(* IEC 61131-3 sources: IRIS-Project/LASAL CONTROL SOFTWARE/LasalProject_2025_09_12/Runtime/%LASALAPPDATA%/Runtime/Library/Loader/Source/code (part 9) *)

END_FUNCTION

//------------------------------------------------------------------------------
// RecvBuf
//
//  This function reads data from a connection. The data is buffered. A tcp-recv
//  operation receives as much data as possible into the internal rx buffer.
//  Data that is not needed by the caller remains in the internal rx buffer.
//  This techniqe is used to avoid multiple small reads from the tcp/ip
//  connection.
//
// Return value
//  If the function succeeds, the return value is the number of bytes read,
//  otherwise a tcp-user error code is returned.
//------------------------------------------------------------------------------
FUNCTION RecvBuf
VAR_INPUT
    bsock         : ^bufferedSocket;
    buf           : ^CHAR;
    len           : UDINT;
    timeout_ms    : UDINT;      // timeout, in milliseconds
END_VAR
VAR_OUTPUT
    retval        : DINT;
END_VAR
VAR
    reqMsg        : msgNopReq;
END_VAR

  #ifdef DEBUG
  ChkBuffer(bsock);
  #endif

  IF bsock^.bytesInRxBuf = 0 THEN
    // The receive buffer is empty

    // Receive as much as possible into the rx buffer
    retval := OS_TCP_USER_RECV(bsock^.sock,
                               #bsock^.rxBuf[0],
                               bsock^.sizeOfRxBuf,
                               0,
                               timeout_ms
                               );
    IF retval <= 0 THEN
#ifdef DEBUG
      IF (retval <> TCP_NOT_READY) | (timeout_ms > 0) THEN
        DEBUGLOG2("%010d-OS_TCP_USER_RECV(sock %d) failed, rc=%d", TO_UDINT(bsock^.sock), TO_UDINT(retval));
      END_IF;
#endif
      IF retval <> TCP_NOT_READY THEN
        CloseBufferedSock(bsock);
      END_IF;
      RETURN;
    END_IF;
    bsock^.bytesInRxBuf += TO_UDINT(retval);
    DEBUG_VERBOSE3("%010d-OS_TCP_USER_RECV(sock %d): %d bytes received, new bytesInRxBuf=%d", TO_UDINT(bsock^.sock), TO_UDINT(retval), TO_UDINT(bsock^.bytesInRxBuf));

    IF bsock^.fAckRcvdData THEN
      // send something after data received to avoid delayed ack
      IF bsock^.bytesInTxBuf > 0 THEN
        FLUSH_TXBUF(bsock);
      ELSE
        SendCmdMsg(bsock,
                   CMD_NOP,
                   0,                 // Type and Ack field of command (type: request, ack: no response is required)
                   #reqMsg$cMessage,
                   SIZEOF(reqMsg),
                   0,                 // timeout: 5 sec.
                   1,                 // use buffered sends
                   1                  // fFlush
                  );
      END_IF;
    END_IF;

  END_IF; // empty rx buffer

  // copy data from the buffer to the caller
  IF len < bsock^.bytesInRxBuf THEN
    retval := len$DINT;
  ELSE
    retval := bsock^.bytesInRxBuf$DINT;
  END_IF;
  IF buf <> NIL THEN
    _memcpy(buf, #bsock^.rxBuf[bsock^.rxBufStrtInd], TO_UDINT(retval));
  END_IF;

  // adjust buffer variables
  bsock^.bytesInRxBuf -= TO_UDINT(retval);
  bsock^.rxBufStrtInd += TO_UDINT(retval);
  IF bsock^.bytesInRxBuf = 0 THEN
    bsock^.rxBufStrtInd := 0;
  END_IF;

  #ifdef DEBUG
  ChkBuffer(bsock);
  #endif

END_FUNCTION

//------------------------------------------------------------------------------
// UnRecvBuf
//
//  This function places len bytes back into the internal rx buffer.
//
// Return value
//  The number of bytes placed into the buffer.
//------------------------------------------------------------------------------
FUNCTION UnRecvBuf
VAR_INPUT
    bsock          : ^bufferedSocket;
    buf            : ^CHAR;
    len            : UDINT;
END_VAR
VAR_OUTPUT
    retval         : UDINT;
END_VAR
VAR
    bytesFree      : UDINT;    // total number of free bytes in the rx buffer
END_VAR

  #ifdef DEBUG
  ChkBuffer(bsock);
  #endif

  bytesFree      := bsock^.sizeOfRxBuf - bsock^.bytesInRxBuf;

  IF len < bytesFree THEN
    retval := len;
  ELSE
    retval := bytesFree;
  END_IF;

  IF retval > bsock^.rxBufStrtInd THEN
    // move the data in rxBuf to the end of the buffer
    _memmove(#bsock^.rxBuf[retval], #bsock^.rxBuf[bsock^.rxBufStrtInd], bsock^.bytesInRxBuf);
    bsock^.rxBufStrtInd := retval;
  END_IF;

  bsock^.rxBufStrtInd -= retval;
  bsock^.bytesInRxBuf += retval;
  _memcpy(#bsock^.rxBuf[bsock^.rxBufStrtInd], buf, retval);

  #ifdef DEBUG
  ChkBuffer(bsock);
  #endif

END_FUNCTION

//------------------------------------------------------------------------------
// ReadN
//
//  This function reads n bytes from a connection.
//
// Return value
//  If the function succeeds, the return value is the number of bytes requested,
//  otherwise a tcp-user error code is returned.
//------------------------------------------------------------------------------
FUNCTION ReadN
VAR_INPUT
    bsock         : ^bufferedSocket;
    buf           : ^CHAR;
    len           : UDINT;
    timeout_ms    : UDINT;      // timeout, in milliseconds
END_VAR
VAR_OUTPUT
    retval        : DINT;
END_VAR
VAR
    ptr           : ^CHAR;
    bytesToRead   : UDINT;      // number of bytes to read
    bytesRead     : UDINT;      // number of bytes already read
END_VAR

    bytesToRead := len;
    bytesRead   := 0;
    ptr         := buf;
    WHILE bytesToRead > 0 DO
      retval := RecvBuf(bsock, ptr, bytesToRead, timeout_ms);
      IF retval <= 0 THEN
        // In the case of an error place already read data back to the buffer
        IF UnRecvBuf(bsock, buf, bytesRead) <> bytesRead THEN
          // This code should never be reached !
          DEBUGLOG1("%010d-ReadN(sock %d): UnRecvBuf failed", TO_UDINT(bsock^.sock));
          CloseBufferedSock(bsock);
          retval := ERR_CONN_BROKEN;
        END_IF;
        RETURN;
      END_IF;
      bytesToRead -= retval$UDINT;
      bytesRead   += retval$UDINT;
      ptr         += retval;
    END_WHILE;

    retval := bytesRead$DINT;

END_FUNCTION

//------------------------------------------------------------------------------
// ReadVRec
//
//  This function reads a record with a variable length.
//
// Return value
//  If the function succeeds, the return value is the number of bytes received
//  in the data field (without vrec-header).
//
// Remarks
//  When the size of the buffer is too small for the message, the connection is
//  closed.
//------------------------------------------------------------------------------
FUNCTION ReadVRec
VAR_INPUT
    bsock         : ^bufferedSocket;
    vrec          : ^vRecord;    // the variable record buffer
    len           : UDINT;      // length of the buffer incl. header
    timeout_ms    : UDINT;      // timeout, in milliseconds
END_VAR
VAR_OUTPUT
    retval        : DINT;
END_VAR

  // first read the vrec-header
  retval := ReadN(bsock, (#vrec^.vHdr)$^CHAR, SIZEOF(vrec^.vHdr), timeout_ms);
  IF retval <= 0 THEN
    RETURN;
  END_IF;

  // check if the header is valid
  IF vrec^.vHdr.id <> 0xFACE THEN
    DEBUGLOG1("%010d-ReadVRec(sock %d): invalid vrec-hdr received", TO_UDINT(bsock^.sock));
    CloseBufferedSock(bsock);
    retval := ERR_INVALID_VRECHDR;
    RETURN;
  END_IF;

  // check how many data fits into the buffer
  IF (vrec^.vHdr.dataLen + SIZEOF(vrec^.vHdr)) > len THEN
    DEBUGLOG1("%010d-ReadVRec(sock %d): buffer too small", TO_UDINT(bsock^.sock));
    CloseBufferedSock(bsock);
    retval := ERR_BUF_TOO_SMALL;
    RETURN;
  END_IF;

  // read the data of the variale record
  retval := ReadN(bsock, (#vrec^.data)$^CHAR, vrec^.vHdr.dataLen, timeout_ms);
  IF retval <= 0 THEN
    // error: write the vrec-header back to the buffer
    IF UnRecvBuf(bsock, (#vrec^.vHdr)$^CHAR, SIZEOF(vrec^.vHdr)) <> SIZEOF(vrec^.vHdr) THEN
      // This code should never be reached !
      DEBUGLOG1("%010d-ReadVRec(sock %d): UnRecvBuf failed", TO_UDINT(bsock^.sock));
      CloseBufferedSock(bsock);
      retval := ERR_CONN_BROKEN;
    END_IF;
    RETURN;
  END_IF;

END_FUNCTION

//------------------------------------------------------------------------------
// ReadCmdMsg
//
//  This function reads a command message.
//
// Return value
//  If the function succeeds, the return value is the number of bytes received
//  in the data field (without vrec-header).
//
// Remarks
//  When the size of the buffer is too small for the message, the rest of the
//  message received and discarded.
//------------------------------------------------------------------------------
FUNCTION ReadCmdMsg
VAR_INPUT
    bsock         : ^bufferedSocket;
    msg           :^cMessage;   // the message
    len           : UDINT;      // length of the message incl. header
    timeout_ms    : UDINT;      // timeout, in milliseconds
    ack           :^UDINT;      // acknowledge field received (optional)
    cmd           : UDINT;      // matching command of the message (n/a for requests)
    typeMask      : UDINT;      // specifies which type (req.,resp.or both) is expected
END_VAR
VAR_OUTPUT
    retval        : DINT;
END_VAR

  retval := ReadVRec(bsock, msg$^vRecord, len, timeout_ms);
  IF retval <= 0 THEN
    RETURN;
  END_IF;

  IF retval < SIZEOF(msg^.cHdr.cmd) THEN
    // at least the header must be available
    DEBUGLOG1("%010d-ReadCmdMsg(sock %d): missing cmd-hdr", TO_UDINT(bsock^.sock));
    CloseBufferedSock(bsock);
    retval := ERR_INVALID_CMSGHDR;
    RETURN;
  END_IF;

  // check if the type of message is expected by the caller
  IF msg^.cHdr.cmd AND MASK_CMD_ISRESP THEN
     // a response is received

    IF (typeMask AND CMD_TYPE_RESP) = 0 THEN
      DEBUGLOG1("%010d-ReadCmdMsg(sock %d): unexpected resonse received", TO_UDINT(bsock^.sock));
      CloseBufferedSock(bsock);
      retval := ERR_INVALID_CMSGTYPE;
    END_IF;
    IF (msg^.cHdr.cmd AND MASK_CMD_CODE) <> cmd THEN
      DEBUGLOG1("%010d-ReadCmdMsg(sock %d): cmd-code in response does not match", TO_UDINT(bsock^.sock));
      CloseBufferedSock(bsock);
      retval := ERR_INVALID_CMSGCODE;
    END_IF;
    IF (msg^.cHdr.cmd AND MASK_CMD_ACK) = 0 THEN
      DEBUGLOG1("%010d-ReadCmdMsg(sock %d): nack received", TO_UDINT(bsock^.sock));
      CloseBufferedSock(bsock);
      retval := ERR_NACK_RECEIVED;
    END_IF;

  ELSE
    // a request is received

    IF (typeMask AND CMD_TYPE_REQ) = 0 THEN
      DEBUGLOG1("%010d-ReadCmdMsg(sock %d): unexpected request received", TO_UDINT(bsock^.sock));
      CloseBufferedSock(bsock);
      retval := ERR_INVALID_CMSGTYPE;
    END_IF;

  END_IF;

  // extract the ack field
  IF ack <> NIL THEN
    ack^ := msg^.cHdr.cmd AND MASK_CMD_ACK;
  END_IF;

END_FUNCTION

//------------------------------------------------------------------------------
// UpdateCell
//
// Return value:
//  Error                                                     : <=0
//  When udLastUpdate did not expire                          : 1
//  When udLastUpdate expired, but dData did not change       : 2
//  When udLastUpdate expired, and dData changed (transfer)   : 3
//------------------------------------------------------------------------------
#ifdef COMLINK_TCP_SERVER
FUNCTION UpdateCell
VAR_INPUT
    pRefrConn     : ^refrConnBlock;
    pUpdCell      : ^comStCell;  // pointer to cell in updatelist
    iOff          : UINT;
END_VAR
VAR_OUTPUT
    retval        : DINT;
END_VAR
VAR
    reqMsg        : msgUpdCellReq; // request structure for command CMD_UPDCELL
    dData         : DINT;
    rc            : DINT;
END_VAR

  retval := 1;

  if( pUpdCell = NIL )then
    return;
  end_if;

  IF pRefrConn^.bsock.fTxBufferShortage <> 0 THEN
    // in the case of a buffer shortage do not send any updatecells
    RETURN;
  END_IF;

  IF QUERY_FREE_TXBUF(pRefrConn^.bsock) < (2 * SIZEOF(reqMsg)) THEN
    // when there is no more space for 2 messages, then enter buffer shortage
    DEBUGLOG0("%010d-UpdateCell: entering tx buffer shortage");
    pRefrConn^.bsock.fTxBufferShortage := 1;
    // try to send all unsent data
    FLUSH_TXBUF(#pRefrConn^.bsock);
  END_IF;

  IF (ops.tAbsolute - pUpdCell^.udLastUpdate) < (pUpdCell^.udUpdateRate AND 16#FFFF) THEN
    // udLastUpdate did not expire
    RETURN;
  END_IF;

  IF pUpdCell^.pCh = NIL THEN
    RETURN;
  END_IF;

  retval := 2;

  IF (pUpdCell^.udUpdateRate and UPDRATE_FLAG_IS_VBI) THEN
    dData := (pUpdCell^.pCh$^virtualBaseInit^.getCrc())$DINT;
  ELSIF (pUpdCell^.udUpdateRate AND UPDRATE_FLAG_IS_MERKEREX) THEN
     dData := (pUpdCell^.pCh$^merkerex^.getcrc())$DINT;
  ELSIF (pUpdCell^.udUpdateRate AND UPDRATE_FLAG_IS_GLOBALVAR) THEN
//    dData := (pUpdCell^.pCh$^DINT)^;
    dData := UpDateGlobalVar(pUpdCell^.pCh, pUpdCell^.udUpdateRate);
  ELSE
    dData := rd(pUpdCell^.pCh);
  END_IF;

  IF dData = pUpdCell^.dData & (pUpdCell^.udUpdateRate and UPDRATE_FLAG_FORCE_CHANGE) = 0 THEN
    // dData did not change
    pUpdCell^.udLastUpdate := ops.tAbsolute;
    RETURN;
  END_IF;
  pUpdCell^.udUpdateRate := pUpdCell^.udUpdateRate AND NOT UPDRATE_FLAG_FORCE_CHANGE;

  retval := 3;

  // prepare the request message structure
  reqMsg.iOff  := iOff;
  reqMsg.pCh   := pUpdCell^.pCh;
  reqMsg.dData := dData;

  // Send the request
  rc := SendCmdMsg(#pRefrConn^.bsock,
                   CMD_UPDCELL,
                   0,                // Type and Ack field of command (type: request, ack: no response required)
                   #reqMsg$cMessage,
                   SIZEOF(reqMsg),
                   0,                // timeout: non-blocking
                   1,                // use buffered sends
                   pRefrConn^.bsock.fTxBufferShortage // fFlush
                  );
  IF rc <= 0 THEN
    DEBUGLOG2("%010d-*** UpdateCell(VarPos %d): SendCmdMsg failed, rc=%d", TO_UDINT(iOff), TO_UDINT(rc));
    retval := rc;
  ELSE
    //DEBUGLOG3("%010d-UpdateCell: UPDCELL request sent, conn=0x%08X, VarPos=%d, dData=0x%08X", pRefrConn$UDINT, TO_UDINT(iOff), TO_UDINT(dData));
    pUpdCell^.dData := dData;
    pUpdCell^.udLastUpdate := ops.tAbsolute;
  END_IF;

END_FUNCTION
#endif

//------------------------------------------------------------------------------
// UpdateListProcessor
//------------------------------------------------------------------------------
#ifdef COMLINK_TCP_SERVER
FUNCTION UpdateListProcessor
VAR_INPUT
    pRefrConn     : ^refrConnBlock;
END_VAR
VAR
    list          : ^updateList;
    pUpdCell      : ^comStCell;  // pointer to cell in updatelist
    pStrtCell     : ^comStCell;
END_VAR

  if( pRefrConn = NIL )then
    return;
  end_if;
  if( pRefrConn^.ptr = NIL )then
    return;
  end_if;
  list := #pRefrConn^.ptr^.statList;
  if( list = NIL )then
    return;
  end_if;

  IF list^.nbrRefrCells > 0 THEN
    pStrtCell := list^.pActCell;
    WHILE 1 DO
      pUpdCell := list^.pActCell;

      UpdateCell(pRefrConn, pUpdCell, list^.actInd$UINT);
      IF pRefrConn^.bsock.sock < 0 THEN
        RETURN;
      END_IF;

      IF (list^.actInd + 1) >= list^.nbrRefrCells THEN
        list^.actInd   := 0;
        list^.pActCell := list^.pFirstCell;
      ELSE
        list^.actInd   += 1;
        list^.pActCell += SIZEOF(list^.pActCell^);
      END_IF;

      IF pStrtCell = list^.pActCell THEN
        EXIT;
      END_IF;
    END_WHILE;
  END_IF;

  list := #pRefrConn^.ptr^.dynList;
  if( list = NIL )then
    return;
  end_if;
  IF list^.nbrRefrCells > 0 THEN
    pStrtCell := list^.pActCell;
    WHILE 1 DO
      pUpdCell := list^.pActCell;

      if( pUpdCell = NIL )then
        return;
      end_if;
      UpdateCell(pRefrConn, pUpdCell, (list^.actInd + 1000)$UINT);
      IF pRefrConn^.bsock.sock < 0 THEN
        RETURN;
      END_IF;

      IF (list^.actInd + 1) >= list^.nbrRefrCells THEN
        list^.actInd   := 0;
        list^.pActCell := list^.pFirstCell;
      ELSE
        list^.actInd   += 1;
        list^.pActCell += SIZEOF(list^.pActCell^);
      END_IF;

      IF pStrtCell = list^.pActCell THEN
        EXIT;
      END_IF;
    END_WHILE;
  END_IF;

END_FUNCTION
#endif

//------------------------------------------------------------------------------
// SendAliveMessage_TCP
//------------------------------------------------------------------------------
#ifdef COMLINK_TCP_SERVER
FUNCTION SendAliveMessage_TCP
VAR_INPUT
    pRefrConn     : ^refrConnBlock;
END_VAR
VAR_OUTPUT
    retval        : DINT;
END_VAR
VAR
    reqMsg        : msgIamAliveReq; // request structure for command CMD_UPDCELL
    rc            : DINT;
END_VAR

  retval := 1;

  IF pRefrConn^.bsock.fTxBufferShortage <> 0 THEN
    // in the case of a buffer shortage do not send any requests
    RETURN;
  END_IF;

  IF QUERY_FREE_TXBUF(pRefrConn^.bsock) < (2 * SIZEOF(reqMsg)) THEN
    // when there is no more space for 2 messages, then enter buffer shortage
    DEBUGLOG0("%010d-SendAliveMessage_TCP: entering tx buffer shortage");
    pRefrConn^.bsock.fTxBufferShortage := 1;
    // try to send all unsent data
    FLUSH_TXBUF(#pRefrConn^.bsock);
  END_IF;

  // Send the request
  rc := SendCmdMsg(#pRefrConn^.bsock,
                   CMD_IAMALIVE,
                   0,                // Type and Ack field of command (type: request, ack: no response required)
                   #reqMsg$cMessage,
                   SIZEOF(reqMsg),
                   0,                // timeout: non-blocking
                   1,                // use buffered sends
                   1                 // fFlush
                  );
  IF rc <= 0 THEN
    DEBUGLOG1("%010d-*** SendAliveMessage_TCP: SendCmdMsg failed, rc=%d", TO_UDINT(rc));
    retval := rc;
  ELSE
    DEBUG_VERBOSE1("%010d-SendAliveMessage_TCP: IAMALIVEL request sent, conn=0x%08X", pRefrConn$UDINT);
  END_IF;
END_FUNCTION
#endif

//------------------------------------------------------------------------------
// SyncRefListsTcp  - siehe Beschreibung von SyncRefLists
//------------------------------------------------------------------------------
#ifdef COMLINK_TCP_SERVER
FUNCTION SyncRefListsTcp
VAR_INPUT
    pCmdConn    : ^cmdConnBlock;
END_VAR
VAR
    obj         : pVoid;
    pHead       : ^IprHead;
    instr       : ^instruct;
    pRefrConn   : ^refrConnBlock;
END_VAR

    pRefrConn := pRefrConnRoot;
    WHILE pRefrConn <> NIL DO
        IF pRefrConn^.ipAddrPeer = pCmdConn^.ipAddrPeer THEN

#ifndef DUMMY_LOADER
            pHead := pCmdConn^.ptr^.com.GetHead();
#endif
            instr := pHead^.pCode;

            IF instr^.opCode = I_WRITE THEN

                obj := instr^.aPara[0]$^pVoid;

                // statische Refresh-Liste durchsuchen
                InvalidateRefListEntry(pRefrConn^.ptr^.statList.pFirstCell, pRefrConn^.ptr^.statList.nbrRefrCells$UINT, obj);

                // dynamische Refresh-Liste durchsuchen
                InvalidateRefListEntry(pRefrConn^.ptr^.dynList.pFirstCell, pRefrConn^.ptr^.dynList.nbrRefrCells$UINT, obj);

            END_IF;

        END_IF;
        pRefrConn := pRefrConn^.next;
    END_WHILE;

END_FUNCTION

FUNCTION GLOBAL SyncRefListsTcpAll
  VAR_INPUT
    lasalid : udint;
  END_VAR
  var
    pRefrConn   : ^refrConnBlock;
  end_var

  pRefrConn := pRefrConnRoot;

  while(pRefrConn <> NIL) do
    // statische Refresh-Liste durchsuchen
    InvalidateRefListEntry(pRefrConn^.ptr^.statList.pFirstCell, pRefrConn^.ptr^.statList.nbrRefrCells$UINT, lasalid$^void);

    // dynamische Refresh-Liste durchsuchen
    InvalidateRefListEntry(pRefrConn^.ptr^.dynList.pFirstCell, pRefrConn^.ptr^.dynList.nbrRefrCells$UINT, lasalid$^void);
    pRefrConn := pRefrConn^.next;
  end_while;

END_FUNCTION
#endif

//------------------------------------------------------------------------------
// Entfernt unbenutzte Verbindungen.
// Es werden alle Verbindungen mit einer bestimmten Remote-IP-Adresse untersucht.
// Wenn die Inst-ID nicht mit der angegebenen übereinstimmt, dann kann es sich
// nur um einen Neustart der Station mit dieser IP-Adresse handeln, da die
// Inst-ID beim Comlink-Init immer neu vergeben wird.
//
// Verbindungen, bei denen die Inst-ID für eine längere Zeit 0 ist, werden
// ebenfalls beendet. Hier handelt es sich um Verbindungen, bei denen abgesteckt
// wurde, bevor CMD_SESSINFO empfangen worden ist.
//
// ApplicationID:
// Wird nur von Comlink Verbindungen von PC-Anwendungen verwendet.
// Wenn auf einem PC mehrere Anwendungen eine Comlink Verbindung verwenden,
// dann kann jede Anwendung eine eigene ApplicationID mitschicken. Damit wird
// verhindert, dass die zweite Anwendung die Verbindung der ersten löscht.
//------------------------------------------------------------------------------
#ifdef COMLINK_TCP_SERVER
FUNCTION DeleteUnusedConnections
VAR_INPUT
    ipAddrPeer   : UDINT;
    instIdOfPeer : UDINT;
    ApplicationID : UDINT;  // ApplicationID
END_VAR
VAR
    pCmdConn   : ^cmdConnBlock;
    pRefrConn   : ^refrConnBlock;
    pCmdConn_next   : ^cmdConnBlock;
    pRefrConn_next  : ^refrConnBlock;
END_VAR

    pCmdConn := pCmdConnRoot;
    WHILE pCmdConn <> NIL DO
        pCmdConn_next := pCmdConn^.next;
        IF ((pCmdConn^.ipAddrPeer = ipAddrPeer) &
            (pCmdConn^.ptr^.instIdOfPeer <> 0) &
            (pCmdConn^.ptr^.instIdOfPeer <> instIdOfPeer) &
            (pCmdConn^.ApplicationID = ApplicationID))
            |
           ((pCmdConn^.ptr^.instIdOfPeer = 0) &
            ((ops.tAbsolute - pCmdConn^.connectTime) > 5000)) THEN
            DEBUGLOG1("%010d-  =====  unused Cmd conn.data block found (ip 08%X) -> releasing block  =====", ipAddrPeer);
            ReleaseConnBlock(TYPE_CMD_CONN, pCmdConn$^connBlock, 0);
            pCmdConn := NIL;
        END_IF;
        pCmdConn := pCmdConn_next;
    END_WHILE;

    pRefrConn := pRefrConnRoot;
    WHILE pRefrConn <> NIL DO
        pRefrConn_next := pRefrConn^.next;
        IF ((pRefrConn^.ipAddrPeer = ipAddrPeer) &
            (pRefrConn^.ptr^.instIdOfPeer <> 0) &
            (pRefrConn^.ptr^.instIdOfPeer <> instIdOfPeer) &
            (pRefrConn^.ApplicationID = ApplicationID))
            |
           ((pRefrConn^.ptr^.instIdOfPeer = 0) &
            ((ops.tAbsolute - pRefrConn^.connectTime) > 5000)) THEN
            DEBUGLOG1("%010d-  =====  unused Refr conn.data block found (ip 08%X) -> releasing block  =====", ipAddrPeer);
            ReleaseConnBlock(TYPE_REFR_CONN, pRefrConn$^connBlock, 0);
            pRefrConn := NIL;
        END_IF;
        pRefrConn := pRefrConn_next;
    END_WHILE;

END_FUNCTION
#endif

//------------------------------------------------------------------------------
// DeleteUnusedRecycleData
//
//  Es werden unbenutzte refresh-connection-data-block's im recycle pool
//  gesucht und wenn gefunden, dann freigegeben.
//
//  Kriterium, ob ein data-block unbenutzt ist:
//  - IP Adresse muss übereinstimmen
//  - InstanceId muss vorhanden, aber unterschiedlich sein
//  - ApplicationID muss übereinstimmen
//------------------------------------------------------------------------------
#ifdef COMLINK_TCP_SERVER
FUNCTION DeleteUnusedRecycleData
VAR_INPUT
    ipAddrPeer   : UDINT;
    instIdOfPeer : UDINT;
    ApplicationID : UDINT;  // ApplicationID
END_VAR
VAR
    pDataWork : ^refrConnData;
    pDataPrev : ^refrConnData;
END_VAR

  pDataPrev := NIL;
  pDataWork := pRefrConnDataRoot;
  WHILE pDataWork <> NIL DO
    IF ((pDataWork^.ipAddrPeer = ipAddrPeer) &
        (pDataWork^.instIdOfPeer <> 0) &
        (pDataWork^.instIdOfPeer <> instIdOfPeer) &
        (pDataWork^.ApplicationID = ApplicationID)) THEN
      // remove it from the recycle pool
      IF pDataPrev = NIL THEN
        pRefrConnDataRoot  := pDataWork^.next;
      ELSE
        pDataPrev^.next := pDataWork^.next;
      END_IF;
      DEBUGLOG1("%010d-  =====  unused recycle refr conn.data block found (ip 08%X) -> releasing block  =====", ipAddrPeer);
      FreeRefrConnData(pDataWork);
      nbrRecycled -= 1;
      EXIT;
    END_IF;
    pDataPrev := pDataWork;
    if( pDataWork = pDataWork^.next )then
      exit;
    end_if;
    pDataWork := pDataWork^.next;
  END_WHILE;

END_FUNCTION
#endif

//------------------------------------------------------------------------------
// CmdMsgListener
//
//  This function serves incoming requests from the client on the command
//  channel.
//------------------------------------------------------------------------------
#ifdef COMLINK_TCP_SERVER
FUNCTION CmdMsgListener
VAR_INPUT
    pCmdConn         : ^cmdConnBlock;
END_VAR
VAR_OUTPUT
    retval    : DINT;
END_VAR
VAR
    cmsg      : cMessage512;
    ackRcvd   : UDINT;        // received ack-field
    ackSend   : UDINT;        // ack-field to send
    dataLen   : UDINT;
    bNext     : UDINT;
    msgLen    : UDINT;
    pResu     : ^results;
    cmd       : UDINT;
    pCmdConnTemp : ^cmdConnBlock;
    rc : DINT;
    releaseFlag : UDINT;
END_VAR

  retval := 0;
  releaseFlag := 0;

  #ifdef LOADER_TCP_MODERATE
    if (pCmdConn^.bsock.isDataAvailable = false) then
      return;
    end_if;
  #endif

  rc := ReadCmdMsg(#pCmdConn^.bsock,
                       #cmsg$cMessage,
                       sizeof(cmsg),
                       0,                   // timeout: 0 means non blocking
                       #ackRcvd,            // received ack field
                       0,                   // matching cmd-code (n/a for requests)
                       CMD_TYPE_REQ         // accept only request types
                      );
  IF rc <= 0 THEN
#ifdef DEBUG
    IF rc <> TCP_NOT_READY THEN
      DEBUGLOG2("%010d-*** CmdMsgListener(sock %d): ReadCmdMsg failed, rc=%d", TO_UDINT(pCmdConn^.bsock.sock), TO_UDINT(rc));
    END_IF;
#endif
    RETURN;
  END_IF;

  retval := 1;

  dataLen := cmsg.cHdr.vHdr.dataLen - SIZEOF(cmsg.cHdr.cmd);
  ackSend := 0; // unsupported command
  msgLen  := SIZEOF(cmsg.cHdr);

  cmd := cmsg.cHdr.cmd AND MASK_CMD_CODE;
  CASE cmd OF

    CMD_BEFIPR:
      DEBUG_VERBOSE2("%010d-CmdMsgListener: sock %d - BEFIPR received, dataLen=%d", TO_UDINT(pCmdConn^.bsock.sock), dataLen$UDINT);
      // req-data:
      //    workState   : iprStates;
      //    instr       : instruct;
      // resp-data:
      //    workState   : iprStates;
      //    resu        : results;

      IF (dataLen < SIZEOF(iprStates)) | ((dataLen - SIZEOF(iprStates)) > SIZEOF(instruct)) THEN
        cmsg$msgBefiprResp.workstate := ERROR;
      ELSE
        // execute befipr
#ifndef DUMMY_LOADER
#ifdef LOADER_4_LASAL2
        _memcpy(pCmdConn^.ptr^.com._m.head.pCode, #cmsg$msgBefiprReq.instr, dataLen - SIZEOF(iprStates));
        pCmdConn^.ptr^.com._m.head.workstate := cmsg$msgBefiprReq.workstate;
        pCmdConn^.ptr^.com._m.head.funkSt    := READY;
        pCmdConn^.ptr^.Com._m.resu.uilng :=0;
#else
        _memcpy(pCmdConn^.ptr^.com.head.pCode, #cmsg$msgBefiprReq.instr, dataLen - SIZEOF(iprStates));
        pCmdConn^.ptr^.com.head.workstate := cmsg$msgBefiprReq.workstate;
        pCmdConn^.ptr^.com.head.funkSt    := READY;
        pCmdConn^.ptr^.Com.resu.uilng :=0;
#endif
        cmsg$msgBefiprResp.workstate := pCmdConn^.ptr^.com.BEFIPR(#bNext);
#endif
        SyncRefListsTcp(pCmdConn);
      END_IF;

      // prepare the response
      ackSend := MASK_CMD_ACK;  // command processed
      msgLen := SIZEOF(cmsg.cHdr) + SIZEOF(iprStates);
      IF cmsg$msgBefiprResp.workstate <> ERROR THEN
#ifndef DUMMY_LOADER
        pResu := pCmdConn^.ptr^.com.GetResult();
#endif
        IF pResu^.uilng <> 16#FFFF THEN
          IF pResu^.uilng <= SIZEOF(cmsg$msgBefiprResp.resu) THEN
            msgLen += pResu^.uilng;
            _memcpy(#cmsg$msgBefiprResp.resu, pResu, pResu^.uilng);
          ELSE
            cmsg$msgBefiprResp.workstate := ERROR;
          END_IF;
        END_IF;
      END_IF;

    CMD_SESSINFO:
      DEBUGLOG2("%010d-CmdMsgListener: sock %d - SESSINFO received, dataLen=%d", TO_UDINT(pCmdConn^.bsock.sock), dataLen$UDINT);
      // req-data:
      //    version     : UDINT;
      // resp-data:
      //    version     : UDINT;

      IF dataLen >= (msgSessInfo.sizeofDynList - msgSessInfo.version) THEN

        pCmdConn^.ApplicationID := 0; // ApplicationID
        IF(datalen >= (msgSessInfo2.ApplicationID - msgSessInfo2.version + 4)) THEN  // ApplicationID
          pCmdConn^.ApplicationID := cmsg$msgSessInfo2.ApplicationID; // ApplicationID
        END_IF; // ApplicationID

        DEBUGLOG3("%010d- instId=%d, appId=%d, sessId=%d", TO_UDINT(cmsg$msgSessInfo.instId), TO_UDINT(pCmdConn^.ApplicationID), TO_UDINT(cmsg$msgSessInfo.sessId));

        // Inaktive Cmd-Connections suchen und freigeben
        pCmdConnTemp := pCmdConnRoot;
        WHILE pCmdConnTemp <> NIL DO

          IF pCmdConnTemp <> pCmdConn THEN
            IF (pCmdConnTemp^.ptr^.instIdOfPeer = cmsg$msgSessInfo.instId) &
               (pCmdConnTemp^.ApplicationID = pCmdConn^.ApplicationID) & // ApplicationID
               (pCmdConnTemp^.ptr^.sessIdOfPeer = cmsg$msgSessInfo.sessId) THEN
               DEBUGLOG0("%010d-  =====  a cmd conn.data block was found in the active list -> releasing block  =====");
               ReleaseConnBlock(TYPE_CMD_CONN, pCmdConnTemp$^connBlock, 0);
               pCmdConnTemp := NIL;
              EXIT;
            END_IF;
          END_IF;

          pCmdConnTemp := pCmdConnTemp^.next;

        END_WHILE;

        // store the information in my context
        pCmdConn^.ptr^.instIdOfPeer := cmsg$msgSessInfo.instId;
        pCmdConn^.ptr^.sessIdOfPeer := cmsg$msgSessInfo.sessId;

        DeleteUnusedConnections(pCmdConn^.ipAddrPeer, pCmdConn^.ptr^.instIdOfPeer, pCmdConn^.ApplicationID);

        // prepare the response
        ackSend := MASK_CMD_ACK;  // command processed
        msgLen := SIZEOF(msgSessInfo);
        cmsg$msgSessInfo.version := COMLINKT_VERSION;
        cmsg$msgSessInfo.instId  := myInstanceID;
        cmsg$msgSessInfo.sessId  := 0;
        cmsg$msgSessInfo.sizeofDynList  := MAX_DYNLIST_ENTRIES;
        cmsg$msgSessInfo.sizeofStatList := MAX_STATLIST_ENTRIES;

#ifdef DEBUG
      ELSE
        DEBUG_VERBOSE0("%010d-CmdMsgListener: dataLen too small");
#endif
      END_IF;

    CMD_LOGOUT:
      DEBUGLOG0("%010d-  =====  LOGOUT CmdConn =====");
      releaseFlag := 1;

    ELSE
      // unknown command
      DEBUGLOG3("%010d-CmdMsgListener: sock %d - unknown command received, cmd=0x%X, dataLen=%d", TO_UDINT(pCmdConn^.bsock.sock), cmd$UDINT, dataLen$UDINT);

  END_CASE;

  IF ackRcvd THEN
    // the received ack field indicates that a response must be sent
    rc := SendCmdMsg(#pCmdConn^.bsock,
                         cmd,
                         MASK_CMD_ISRESP OR MASK_CMD_ACK,  // Type and Ack field of command (type: response, ack: command processed)
                         #cmsg$cMessage,
                         msgLen,          // length of the message incl. header
                         0,               // timeout_ms: no-blocking
                         1,               // useBuffer
                         1                // fFlush
                        );
    IF rc <= 0 THEN
      DEBUGLOG2("%010d-*** CmdMsgListener(sock %d): SendCmdMsg failed, rc=%d", TO_UDINT(pCmdConn^.bsock.sock), TO_UDINT(rc));
      CloseBufferedSock(#pCmdConn^.bsock);
      IF releaseFlag THEN
        ReleaseConnBlock( TYPE_CMD_CONN, pCmdConn$^connBlock, 0 );
        pCmdConn := NIL;
        retval := -1; // zeigt an, dass der Block freigegeben wurde und nicht mehr benutzt werden darf
      END_IF;
      RETURN;
#ifdef DEBUG
    ELSE
      DEBUG_VERBOSE2("%010d-CmdMsgListener: sock %d - cmd response sent, msgLen=%d", TO_UDINT(pCmdConn^.bsock.sock), msgLen$UDINT);
#endif
    END_IF;
  END_IF;

  IF releaseFlag & pCmdConn THEN
    ReleaseConnBlock( TYPE_CMD_CONN, pCmdConn$^connBlock, 0 );
    pCmdConn := NIL;
    retval := -1; // zeigt an, dass der Block freigegeben wurde und nicht mehr benutzt werden darf
  END_IF;

END_FUNCTION
#endif

//------------------------------------------------------------------------------
// RefrMsgListener
//
//  This function serves incoming requests from the client on the refresh
//  channel.
//
// Return value
//  This function returns 0 when no message was received, otherwise a value
//  greater than 0 is returned.
//------------------------------------------------------------------------------
#ifdef COMLINK_TCP_SERVER
FUNCTION RefrMsgListener
VAR_INPUT
    pRefrConn         : ^refrConnBlock;
END_VAR
VAR_OUTPUT
    retval    : DINT;
END_VAR
VAR
    cmsg      : cMessage512;
    ackRcvd   : UDINT;        // received ack-field
    ackSend   : UDINT;        // ack-field to send
    dataLen   : UDINT;
    msgLen    : UDINT;
    cmd       : UDINT;
    updList   : ^updateList;
    listType  : UDINT;
    pComCell  : ^comStCell;
    udLastUpdate : UDINT;
    pData     : ^refrConnData;
    pRefrConnTemp : ^refrConnBlock;
    rc        : DINT;
    releaseFlag : UDINT;
END_VAR

  retval := 0;
  releaseFlag := 0;

  #ifdef LOADER_TCP_MODERATE
    if (pRefrConn^.bsock.isDataAvailable = false) then
      return;
    end_if;
  #endif

  rc := ReadCmdMsg(#pRefrConn^.bsock,
                   #cmsg$cMessage,
                   SIZEOF(cmsg),
                   0,                   // timeout: 0 means non blocking
                   #ackRcvd,            // received ack field
                   0,                   // matching cmd-code (n/a for requests)
                   CMD_TYPE_REQ         // accept only request types
                  );
  IF rc <= 0 THEN
#ifdef DEBUG
    IF rc <> TCP_NOT_READY THEN
      DEBUGLOG2("%010d-*** RefrMsgListener(sock %d): ReadCmdMsg failed, rc=%d", pRefrConn^.bsock.sock$UDINT, TO_UDINT(rc));
    END_IF;
#endif
    #ifdef LOADER_TCP_MODERATE
      pRefrConn^.bsock.isDataAvailable := false;
    #endif
    RETURN;
  END_IF;

  retval := 1;

  dataLen := cmsg.cHdr.vHdr.dataLen - SIZEOF(cmsg.cHdr.cmd);
  ackSend := 0; // unsupported command
  msgLen  := SIZEOF(cmsg.cHdr);

  cmd := cmsg.cHdr.cmd AND MASK_CMD_CODE;
  CASE cmd OF

    CMD_TXUPD:
      DEBUG_VERBOSE3("%010d-RefrMsgListener: sock %d - TXUPD received, dataLen=%d, VarPos=%d", pRefrConn^.bsock.sock$UDINT, dataLen$UDINT, TO_UDINT(cmsg$msgTxUpdReq.iOff));
      // req-data:
      //    iOff        : UINT;
      //    comcell     : comStCell;
      // resp-data:
      //    this request requires no response

      IF dataLen >= (SIZEOF(msgTxUpdReq) - SIZEOF(msgTxUpdReq.cHdr)) THEN
        IF cmsg$msgTxUpdReq.iOff < 1000 THEN
          updList   := #pRefrConn^.ptr^.statList;
          listType  := 0;
        ELSE
          updList   := #pRefrConn^.ptr^.dynList;
          listType  := 1;
          cmsg$msgTxUpdReq.iOff -=1000;
        END_IF;

        if( updList^.pFirstCell = NIL )then
          return;
        end_if;

        IF TO_UDINT(cmsg$msgTxUpdReq.iOff) >= updList^.nbrCells THEN
          IF IncreaseUpdateList(updList, TO_UDINT(cmsg$msgTxUpdReq.iOff) + 1, listType) = NIL THEN
            DEBUGLOG1("%010d-*** RefrMsgListener: sock %d - MemoryUpdateList failed", pRefrConn^.bsock.sock$UDINT);
            CloseBufferedSock(#pRefrConn^.bsock);
            RETURN;
          END_IF;
          DEBUGLOG3("%010d-*** RefrMsgListener: sock %d - updList %d increased to %d entries", pRefrConn^.bsock.sock$UDINT, listType, updList^.nbrCells);
        END_IF;

        pComCell := updList^.pFirstCell + (SIZEOF(comStCell) * cmsg$msgTxUpdReq.iOff);

        IF (cmsg$msgTxUpdReq.comcell.pCh <> pComCell^.pCh) |
           ((cmsg$msgTxUpdReq.comcell.udUpdateRate AND 0xF0000000) <> (pComCell^.udUpdateRate AND 0xF0000000)) |
           (cmsg$msgTxUpdReq.iOff >= updList^.nbrRefrCells) THEN
          // Es handelt sich um eine geänderte oder neue Zelle
          // -> Werte so setzen, damit gleich einmal ein Refresh passiert
          DEBUGLOG1("%010d-CMD_TXUPD: new cell %d", TO_UDINT(cmsg$msgTxUpdReq.iOff));
          pComCell^ := cmsg$msgTxUpdReq.comcell;
          pComCell^.dData        := 16#80000001$DINT; // invalid
          pComCell^.udUpdateRate := pComCell^.udUpdateRate or UPDRATE_FLAG_FORCE_CHANGE;
          pComCell^.udLastUpdate := ops.tAbsolute - 20*60*1000;  // current time - 20min.
        ELSE
          // Die Zelle hat es schon gegeben. udLastUpdate wird nicht geändert, da kein
          // Refresh notwendig ist
          DEBUGLOG1("%010d-CMD_TXUPD: re-used cell %d", TO_UDINT(cmsg$msgTxUpdReq.iOff));
          udLastUpdate := pComCell^.udLastUpdate;
          pComCell^ := cmsg$msgTxUpdReq.comcell;
          pComCell^.udLastUpdate := udLastUpdate;
        END_IF;

        IF (pComCell^.udUpdateRate AND 0xFFFF) < SMALLEST_UPD_INTERVALL THEN
          pComCell^.udUpdateRate := (pComCell^.udUpdateRate AND 0xFFFF0000) OR SMALLEST_UPD_INTERVALL;
        END_IF;
        IF !!(pComCell^.udUpdateRate AND UPDRATE_FLAG_IS_GLOBALVAR) &
           GetdataBufferFlag(pComCell^.pCh$^VirtualBase) THEN
          // The object has the flag ATTR_DATA_BUFFER set. For these object more than
          // the 4 bytes of dData can be transmitted. The comlink server updates the cell
          // when the crc changes instead of dData.
          pComCell^.udUpdateRate := pComCell^.udUpdateRate or UPDRATE_FLAG_IS_VBI;
        END_IF;
#ifdef DEBUG
      ELSE
        DEBUG_VERBOSE0("%010d-RefrMsgListener: dataLen too small");
#endif
      END_IF;

    CMD_SSREFR:
      DEBUG_VERBOSE3("%010d-RefrMsgListener: sock %d - SSREFR received, typ=%d, count=%d", pRefrConn^.bsock.sock$UDINT, TO_UDINT(cmsg$msgSsRefrReq.typ), TO_UDINT(cmsg$msgSsRefrReq.count));
      // req-data:
      //    count       : UINT;
      //    typ         : UINT;
      // resp-data:
      //    this request requires no response

      IF dataLen >= (SIZEOF(msgSsRefrReq) - SIZEOF(msgSsRefrReq.cHdr)) THEN
        IF cmsg$msgSsRefrReq.typ = 0 THEN
          // static list
          LoadUpdateList(#pRefrConn^.ptr^.statList, cmsg$msgSsRefrReq.count);
        ELSE
          // dynamic list
          LoadUpdateList(#pRefrConn^.ptr^.dynList, cmsg$msgSsRefrReq.count);
        END_IF;
        // Wenn ein StartStopRefresh empfangen wurde, wird ein Flag gesetzt, das bewirkt,
        // dass die Sends der Abarbeitung der Refreshliste nicht gepuffert sondern gleich
        // gesendet werden.
        pRefrConn^.flushNextSends := TRUE;
#ifdef DEBUG
      ELSE
        DEBUG_VERBOSE0("%010d-RefrMsgListener: dataLen too small");
#endif
      END_IF;

    CMD_NOP:
      DEBUG_VERBOSE1("%010d-RefrMsgListener: sock %d - NOP received", pRefrConn^.bsock.sock$UDINT);
      // req-data:
      //    this request contains not data
      // resp-data:
      //    this request requires no response

    CMD_SESSINFO:
      DEBUGLOG2("%010d-RefrMsgListener: sock %d - SESSINFO received, dataLen=%d", TO_UDINT(pRefrConn^.bsock.sock), dataLen$UDINT);
      // req-data:
      //    version     : UDINT;
      // resp-data:
      //    version     : UDINT;

      IF dataLen >= (msgSessInfo.sizeofDynList - msgSessInfo.version) THEN

        pRefrConn^.ApplicationID := 0; // ApplicationID
        IF(datalen >= (msgSessInfo2.ApplicationID - msgSessInfo2.version + 4)) THEN  // ApplicationID
          pRefrConn^.ApplicationID := cmsg$msgSessInfo2.ApplicationID; // ApplicationID
        END_IF; // ApplicationID

        // Search in all other connections for the same inst-ID and sess-ID.
        // When found, we assume that this is an inactive connection and we close
        // this connection.

        DEBUGLOG3("%010d- instId=%d, appId=%d, sessId=%d", TO_UDINT(cmsg$msgSessInfo.instId), TO_UDINT(pRefrConn^.ApplicationID), TO_UDINT(cmsg$msgSessInfo.sessId));

        // Inaktive Refr-Connections suchen und freigeben
        pRefrConnTemp := pRefrConnRoot;
        WHILE pRefrConnTemp <> NIL DO

          IF pRefrConnTemp <> pRefrConn THEN
            IF (pRefrConnTemp^.ptr^.instIdOfPeer = cmsg$msgSessInfo.instId) &
               (pRefrConnTemp^.ApplicationID = pRefrConn^.ApplicationID) & // ApplicationID
               (pRefrConnTemp^.ptr^.sessIdOfPeer = cmsg$msgSessInfo.sessId) THEN
               DEBUGLOG0("%010d-  =====  a refr.conn.data block was found in the active list -> releasing block  =====");
               ReleaseConnBlock(TYPE_REFR_CONN, pRefrConnTemp$^connBlock, 0);
               pRefrConnTemp := NIL;
              EXIT;
            END_IF;
          END_IF;

          pRefrConnTemp := pRefrConnTemp^.next;

        END_WHILE;

        // Check if we can replace an untouched refresh connection data block
        // with a data block from the recycle pool for reconnect of a client.
        pData := NIL;
        IF pRefrConn^.ptr^.instIdOfPeer = 0 THEN
          // the current refresh connection data block is unused
          pData := ReuseRefrConnData(cmsg$msgSessInfo.instId, cmsg$msgSessInfo.sessId);
          IF pData <> NIL THEN
            // a data block was found in the recycle pool
            // -> free the current data block and use the block from the pool
            DEBUGLOG0("%010d-  =====  re-using connnection data block from a previous connection  =====");
            FreeRefrConnData(pRefrConn^.ptr);
            pRefrConn^.ptr := pData;
            DEBUGLOG2("%010d- statList, nbrCells=%d, nbrRefrCells=%d", pRefrConn^.ptr^.statList.nbrCells, pRefrConn^.ptr^.statList.nbrRefrCells);
            DEBUGLOG2("%010d- dynList,  nbrCells=%d, nbrRefrCells=%d", pRefrConn^.ptr^.dynList.nbrCells,  pRefrConn^.ptr^.dynList.nbrRefrCells);
#ifdef DEBUG
          ELSE
            DEBUGLOG0("%010d-  =====  could not re-use connnection data block from a previous connection  =====");
#endif
          END_IF;
#ifdef DEBUG
        ELSE
          DEBUGLOG0("%010d-  =====  did not try to re-use connnection data block from a previous connection  =====");
#endif
        END_IF;

        // store the information in my context
        pRefrConn^.ptr^.instIdOfPeer := cmsg$msgSessInfo.instId;
        pRefrConn^.ptr^.sessIdOfPeer := cmsg$msgSessInfo.sessId;
        pRefrConn^.ptr^.ipAddrPeer := pRefrConn^.ipAddrPeer;
        pRefrConn^.ptr^.ApplicationID := pRefrConn^.ApplicationID;

        DeleteUnusedConnections(pRefrConn^.ipAddrPeer, pRefrConn^.ptr^.instIdOfPeer, pRefrConn^.ApplicationID);
        DeleteUnusedRecycleData(pRefrConn^.ipAddrPeer, pRefrConn^.ptr^.instIdOfPeer, pRefrConn^.ApplicationID);

        // prepare the response
        ackSend := MASK_CMD_ACK;  // command processed
        msgLen := SIZEOF(msgSessInfo);
        cmsg$msgSessInfo.version := COMLINKT_VERSION;
        cmsg$msgSessInfo.instId  := myInstanceID;
        cmsg$msgSessInfo.sessId  := 0;
        cmsg$msgSessInfo.sizeofDynList  := MAX_DYNLIST_ENTRIES;
        cmsg$msgSessInfo.sizeofStatList := MAX_STATLIST_ENTRIES;

#ifdef DEBUG
      ELSE
        DEBUG_VERBOSE0("%010d-RefrMsgListener: dataLen too small");
#endif
      END_IF;

    CMD_MAXIDLETIME:
      DEBUG_VERBOSE2("%010d-RefrMsgListener: sock %d - CMD_MAXIDLETIME received, maxIdleTime=%d", pRefrConn^.bsock.sock$UDINT, cmsg$msgIdlTimReq.maxIdleTime_ms);
      // req-data:
      //    maxIdleTime_ms : UDINT;
      // resp-data:
      //    this request requires no response

      IF cmsg$msgIdlTimReq.maxIdleTime_ms <> pRefrConn^.ptr^.maxIdleTime_ms THEN
        pRefrConn^.ptr^.maxIdleTime_ms := cmsg$msgIdlTimReq.maxIdleTime_ms;
        pRefrConn^.ptr^.lastSendTime_ms := ops.tAbsolute - pRefrConn^.ptr^.maxIdleTime_ms; // damit gleich was geschickt wird
      END_IF;

    CMD_LOGOUT:
      DEBUG_VERBOSE3("%010d-RefrMsgListener: sock %d - LOGOUT received, typ=%d, count=%d", pRefrConn^.bsock.sock$UDINT, TO_UDINT(cmsg$msgSsRefrReq.typ), TO_UDINT(cmsg$msgSsRefrReq.count));
      // req-data:
      //    this request requires no data
      // resp-data:
      //    this request requires no response
      LoadUpdateList( #pRefrConn^.ptr^.statList, 0 );
      LoadUpdateList( #pRefrConn^.ptr^.dynList, 0 );

      DEBUGLOG0("%010d-  =====  LOGOUT RefrConn  =====");
      releaseFlag := 1;

    ELSE
      // unknown command
      DEBUGLOG2("%010d-RefrMsgListener: sock %d - unknown command received, dataLen=%d", pRefrConn^.bsock.sock$UDINT, dataLen$UDINT);

  END_CASE;

  IF ackRcvd THEN
    // the received ack field indicates that a response must be sent
    rc := SendCmdMsg(#pRefrConn^.bsock,
                     cmd,
                     MASK_CMD_ISRESP OR MASK_CMD_ACK,  // Type and Ack field of command (type: response, ack: command processed)
                     #cmsg$cMessage,
                     msgLen,          // length of the message incl. header
                     0,               // timeout_ms: no-blocking
                     1,               // useBuffer
                     1                // fFlush
                    );
    IF rc <= 0 THEN
      DEBUGLOG2("%010d-*** RefrMsgListener(sock %d): SendCmdMsg failed, rc=%d", TO_UDINT(pRefrConn^.bsock.sock), TO_UDINT(rc));
      IF rc = ERR_BUFFER_SHORTAGE THEN
        LDR_DebugLog0("%010d comlink: closing refr-sock due to buffer shortage");
        _onlineDiagFlags := _onlineDiagFlags OR 2;
      END_IF;
      CloseBufferedSock(#pRefrConn^.bsock);
      IF releaseFlag THEN
        ReleaseConnBlock( TYPE_REFR_CONN, s_pRefrConn$^connBlock, 0 );
        s_pRefrConn := NIL;
        retval := -1; // zeigt an, dass der Block freigegeben wurde und nicht mehr benutzt werden darf
      END_IF;
      RETURN;
#ifdef DEBUG
    ELSE
      DEBUG_VERBOSE2("%010d-RefrMsgListener: sock %d - cmd response sent, msgLen=%d", TO_UDINT(pRefrConn^.bsock.sock), rc$UDINT);
#endif
    END_IF;
  END_IF;

  IF releaseFlag & s_pRefrConn THEN
    ReleaseConnBlock( TYPE_REFR_CONN, s_pRefrConn$^connBlock, 0 );
    s_pRefrConn := NIL;
    retval := -1; // zeigt an, dass der Block freigegeben wurde und nicht mehr benutzt werden darf
  END_IF;

END_FUNCTION
#endif

//------------------------------------------------------------------------------
// AliveCheckMsgRcvd
//------------------------------------------------------------------------------
FUNCTION AliveCheckMsgRcvd
VAR_INPUT
  pLogin         : ^loginContext; // connection context
END_VAR
VAR
	pNode 						  : ^MonitorNode;
END_VAR

    OS_MT_WAIT(monitorNodeMutex);
    pNode := pLogin^.pNode;
    IF pNode THEN
        pNode^.lastRcvdTime_ms := ops.tAbsolute;
        pNode^.isRemotePlcAlive := TRUE;
    END_IF;
    OS_MT_SIGNAL(monitorNodeMutex);

END_FUNCTION

//------------------------------------------------------------------------------
// UpdCellListener
//
//  This function serves incoming requests from the server on the refresh
//  channel.
//
// Return value
//  This function returns 0 when no message was received, otherwise a value
//  greater than 0 is returned.
//------------------------------------------------------------------------------
#ifdef COMLINK_TCP_CLIENT
FUNCTION UpdCellListener
VAR_INPUT
    pLogin         : ^loginContext; // connection context
END_VAR
VAR_OUTPUT
    retval         : UDINT;
END_VAR
VAR
    cmsg      : cMessage512;
    ackRcvd   : UDINT;        // received ack-field
    ackSend   : UDINT;        // ack-field to send
    dataLen   : UDINT;
    msgLen    : UDINT;
    cmd       : UDINT;
    pComCell  : ^comStCell;
    data2LSE  : d2LSE;
    uiOffs    : UINT;
    rc        : DINT;
    original_this : UDINT;
    pCallbackListEntry :^sDynCallbackList;
END_VAR

  retval := 0;

  #ifdef LOADER_TCP_MODERATE
    if (pLogin^.refrSockClnt.isDataAvailable = FALSE) then
      return;
    end_if;
  #endif

  pLogin^.refrSockClnt.fAckRcvdData := 1;

  rc := ReadCmdMsg(#pLogin^.refrSockClnt,
                   #cmsg$cMessage,
                   SIZEOF(cmsg),
                   0,                   // timeout: 0 means non blocking
                   #ackRcvd,            // received ack field
                   0,                   // matching cmd-code (n/a for requests)
                   CMD_TYPE_REQ         // accept only request types
                  );
  IF rc <= 0 THEN
    IF rc <> TCP_NOT_READY THEN
      DEBUGLOG2("%010d-*** UpdCellListener: ReadCmdMsg failed, rc=%d, closing refr sock %d", TO_UDINT(rc), pLogin^.refrSockClnt.sock$UDINT);
      CloseBufferedSock(#pLogin^.refrSockClnt);
    END_IF;
    #ifdef LOADER_TCP_MODERATE
      pLogin^.refrSockClnt.isDataAvailable := false;
    #endif
    RETURN;
  END_IF;
  pLogin^.refrSockClnt.fAckRcvdData := 0;
  AliveCheckMsgRcvd(pLogin);

  retval := 1;

  dataLen := cmsg.cHdr.vHdr.dataLen - SIZEOF(cmsg.cHdr.cmd);
  ackSend := 0; // value for an unsupported command (=nack)
  msgLen  := SIZEOF(cmsg.cHdr);

  cmd := cmsg.cHdr.cmd AND MASK_CMD_CODE;
  CASE cmd OF

    CMD_UPDCELL:
      DEBUG_VERBOSE3("%010d-UpdCellListener: sock %d - UPDCELL received, dataLen=%d, VarPos=%d", pLogin^.refrSockClnt.sock$UDINT, dataLen$UDINT, TO_UDINT(cmsg$msgUpdCellReq.iOff));
      // req-data:
      //    iOff        : INT;
      //    comcell     : comStCell;
      // resp-data:
      //    this request requires no response

      IF dataLen >= (SIZEOF(msgUpdCellReq) - SIZEOF(msgUpdCellReq.cHdr)) THEN
        uiOffs := cmsg$msgUpdCellReq.iOff$UINT;
        IF uiOffs < 1000 THEN
          pComCell := pLogin^.statList.pFirstCell;
          IF TO_UDINT(cmsg$msgUpdCellReq.iOff) >= pLogin^.statList.nbrCells THEN
            DEBUGLOG2("%010d-*** UpdCellListener: sock %d - VarPos(%d) is too big for StatList", pLogin^.refrSockClnt.sock$UDINT, TO_UDINT(cmsg$msgUpdCellReq.iOff));
            RETURN;
          END_IF;
        ELSE
          uiOffs -=1000;
          pComCell := pLogin^.dynlist.pFirstCell;
          IF TO_UDINT(uiOffs) >= pLogin^.dynList.nbrCells THEN
            DEBUGLOG2("%010d-*** UpdCellListener: sock %d - VarPos(%d) is too big for DynList", pLogin^.refrSockClnt.sock$UDINT, TO_UDINT(cmsg$msgUpdCellReq.iOff));
            RETURN;
          END_IF;
        END_IF;

        pComCell        := pComcell + (SIZEOF(comStCell) * uiOffs);

        IF pComCell^.pCh <> cmsg$msgUpdCellReq.pCh THEN
          DEBUGLOG1("%010d-*** UpdCellListener: sock %d - invalid upd-cell received", pLogin^.refrSockClnt.sock$UDINT);
          RETURN;
        END_IF;
        pComCell^.dData := cmsg$msgUpdCellReq.dData;

        // call callback function
        IF ((pLogin^.pCallback <> NIL) | (pLogin^.pDynCallbacks <> NIL)) THEN
          data2LSE.data      := pComCell^.dData;
          data2LSE.uiOffs    := cmsg$msgUpdCellReq.iOff$UINT;
          data2LSE.varlistID := pComCell^.VarlistID;
          original_this := ESI;

          IF (pLogin^.pCallback <> NIL) THEN
             ESI := pLogin^.pThis;
            pLogin^.pCallback$PrototypeCallbackT(pLogin^.pComdefT, #data2LSE);
          END_IF;
          IF (pLogin^.pDynCallbacks <> NIL) THEN
             pCallbackListEntry := pLogin^.pDynCallbacks;
             WHILE ((pCallbackListEntry <> NIL) & (pCallbackListEntry^.pCallback <> NIL)) DO
                ESI := pCallbackListEntry^.pCallback^.pThis;
                pCallbackListEntry^.pCallback^.pCallback$PrototypeCallbackT(pLogin^.pComdefT, #data2LSE);
                pCallbackListEntry := pCallbackListEntry^.pNext;
             END_WHILE;
          END_IF;

          ESI := original_this;

          DEBUG_VERBOSE3("%010d-UpdCellListener: Callback(dData=0x%08X,uiOffs=%d,id=0x%08X", TO_UDINT(data2LSE.data), TO_UDINT(data2LSE.uiOffs), TO_UDINT(data2LSE.varlistID));
        END_IF;

#ifdef DEBUG
      ELSE
        DEBUG_VERBOSE0("%010d-UpdCellListener: dataLen too small");
#endif
      END_IF;

    CMD_IAMALIVE:
      DEBUG_VERBOSE1("%010d-UpdCellListener: sock %d - IAMALIVE received", pLogin^.refrSockClnt.sock$UDINT);
      // req-data:
      // resp-data:
      //    this request requires no response

    ELSE
      // unknown command
      DEBUGLOG2("%010d-UpdCellListener: sock %d - unknown command received, dataLen=%d", pLogin^.refrSockClnt.sock$UDINT, dataLen$UDINT);

  END_CASE;

  IF ackRcvd THEN
    // the received ack field indicates that a response must be sent
    rc := SendCmdMsg(#pLogin^.refrSockClnt,
                     cmd,
                     MASK_CMD_ISRESP OR MASK_CMD_ACK,  // Type and Ack field of command (type: response, ack: command processed)
                     #cmsg$cMessage,
                     msgLen,          // length of the message incl. header
                     0,               // timeout_ms: no-blocking
                     1,               // useBuffer
                     1                // fFlush
                    );
    IF rc <= 0 THEN
      DEBUGLOG2("%010d-*** UpdCellListener: SendCmdMsg failed, rc=%d, closing refr sock %d", TO_UDINT(rc), pLogin^.refrSockClnt.sock$UDINT);
      CloseBufferedSock(#pLogin^.refrSockClnt);
      RETURN;
#ifdef DEBUG
    ELSE
      DEBUG_VERBOSE2("%010d-UpdCellListener: sock %d - cmd response sent, msgLen=%d", TO_UDINT(pLogin^.refrSockClnt.sock), rc$UDINT);
#endif
    END_IF;
  END_IF;

END_FUNCTION
#endif

//------------------------------------------------------------------------------
// PndConnListener
//
//  This function listens on the pending socket for a response of a SESSINFO
//  command.
//------------------------------------------------------------------------------
#ifdef COMLINK_TCP_CLIENT
FUNCTION PndConnListener
VAR_INPUT
    pLogin         : ^loginContext; // connection context
END_VAR
VAR_OUTPUT
    retval         : UDINT;
END_VAR
VAR
    cmsg      : cMessage512;
    ackRcvd   : UDINT;        // received ack-field
    ackSend   : UDINT;        // ack-field to send
    dataLen   : UDINT;
    msgLen    : UDINT;
    cmd       : UDINT;
    rc        : DINT;
END_VAR

  retval := 0;
  IF pLogin^.refrSockClnt.sock < 0 THEN
    RETURN;
  END_IF;

  rc := ReadCmdMsg(#pLogin^.refrSockClnt,
                   #cmsg$cMessage,
                   SIZEOF(cmsg),
                   0,                   // timeout: 0 means non blocking
                   #ackRcvd,            // received ack field
                   0,                   // matching cmd-code (n/a for requests)
                   CMD_TYPE_RESP        // accept only request types
                  );
  IF rc <= 0 THEN
    IF rc <> TCP_NOT_READY THEN
      DEBUGLOG2("%010d-*** PndConnListener: ReadCmdMsg failed, rc=%d, closing refr sock %d", TO_UDINT(rc), pLogin^.refrSockClnt.sock$UDINT);
      CloseBufferedSock(#pLogin^.refrSockClnt);
    END_IF;
    RETURN;
  END_IF;
  AliveCheckMsgRcvd(pLogin);

  retval := 1;

  dataLen := cmsg.cHdr.vHdr.dataLen - SIZEOF(cmsg.cHdr.cmd);
  ackSend := 0; // value for an unsupported command (=nack)
  msgLen  := SIZEOF(cmsg.cHdr);

  cmd := cmsg.cHdr.cmd AND MASK_CMD_CODE;
  CASE cmd OF

    CMD_SESSINFO:
      IF cmsg.cHdr.cmd AND MASK_CMD_ISRESP THEN
        DEBUGLOG2("%010d-PndConnListener: sock %d - SESSINFO response received, dataLen=%d", TO_UDINT(pLogin^.refrSockClnt.sock), dataLen$UDINT);
        // req-data:
        //    version     : UDINT;
        // resp-data:
        //    version     : UDINT;

        IF dataLen >= (msgSessInfo.sizeofDynList - msgSessInfo.version) THEN

          IF pLogin^.refrSockClnt.isInstIdVerified = INSTID_CMD_PENDING THEN
            IF pLogin^.instIdOfPeer = cmsg$msgSessInfo.instId THEN
              DEBUGLOG0("%010d-*** PndConnListener: instance ID matches");
              pLogin^.refrSockClnt.isInstIdVerified := INSTID_MATCH;
            ELSE
              DEBUGLOG0("%010d-*** PndConnListener: instance ID does not match, closeing connection");
              pLogin^.refrSockClnt.isInstIdVerified := INSTID_MISMATCH;
              CloseBufferedSock(#pLogin^.refrSockClnt);
            END_IF;
          END_IF;

#ifdef DEBUG
        ELSE
          DEBUG_VERBOSE0("%010d-PndConnListener: dataLen too small");
#endif
        END_IF;

        IF dataLen >= (msgSessInfo.sizeofStatList + sizeof(msgSessInfo.sizeofStatList) - msgSessInfo.version) THEN
            pLogin^.sizeofRemoteDynList  := cmsg$msgSessInfo.sizeofDynList;
            pLogin^.sizeofRemoteStatList := cmsg$msgSessInfo.sizeofStatList;
        END_IF;

      END_IF;

    ELSE
      // unknown command
      DEBUGLOG2("%010d-PndConnListener: sock %d - unknown command received, dataLen=%d", pLogin^.refrSockClnt.sock$UDINT, dataLen$UDINT);

  END_CASE;

END_FUNCTION
#endif

//------------------------------------------------------------------------------
// SendSessionInfo
//------------------------------------------------------------------------------
#ifdef COMLINK_TCP_CLIENT
FUNCTION SendSessionInfo
VAR_INPUT
    bsock         : ^bufferedSocket;
    mySessId      : UDINT;
    timeout_ms    : UDINT;      // timeout, in milliseconds
END_VAR
VAR_OUTPUT
    retval        : DINT;
END_VAR
VAR
    cmsg          : cMessage256;
    useBuffer     : UDINT;
    fFlush        : UDINT;
END_VAR

  // Send the request
  cmsg$msgSessInfo2.version := COMLINKT_VERSION;
  cmsg$msgSessInfo2.instId  := myInstanceId;
  cmsg$msgSessInfo2.sessId  := mySessId;
  cmsg$msgSessInfo2.sizeofDynList  := MAX_DYNLIST_ENTRIES;
  cmsg$msgSessInfo2.sizeofStatList := MAX_STATLIST_ENTRIES;
  cmsg$msgSessInfo2.applicationId := myApplId;

  IF timeout_ms = 0 THEN
    useBuffer := 1;
    fFlush    := 1;
  ELSE
    useBuffer := 0;
    fFlush    := 0;
  END_IF;

  retval := SendCmdMsg(bsock,
                       CMD_SESSINFO,
                       MASK_CMD_ACK,      // Type and Ack field of command (type: request, ack: a response is required)
                       #cmsg$cMessage,
                       SIZEOF(msgSessInfo2),
                       timeout_ms,
                       useBuffer,
                       fFlush
                      );
  IF retval <= 0 THEN
    DEBUGLOG1("%010d-*** SendSessionInfo: SendCmdMsg(CMD_SESSINFO) failed, retval=%d", TO_UDINT(retval));
    RETURN;
  END_IF;
  DEBUGLOG0("%010d-SendSessionInfo: SESSINFO request sent");

END_FUNCTION
#endif

//------------------------------------------------------------------------------
// RecvSessionInfo
//------------------------------------------------------------------------------
#ifdef COMLINK_TCP_CLIENT
FUNCTION RecvSessionInfo
VAR_INPUT
    bsock         : ^bufferedSocket;
    timeout_ms    : UDINT;      // timeout, in milliseconds
    versionOfPeer : ^UDINT;
    instIdOfPeer  : ^UDINT;
    sizeofRemoteDynList  : ^UINT;
    sizeofRemoteStatList : ^UINT;
END_VAR
VAR_OUTPUT
    retval        : DINT;
END_VAR
VAR
    cmsg          : cMessage256;
END_VAR

  // Read the response
  retval := ReadCmdMsg(bsock,
                       #cmsg$cMessage,
                       SIZEOF(cmsg),
                       timeout_ms,
                       NIL,                 // received ack field
                       CMD_SESSINFO,
                       CMD_TYPE_RESP        // accept only response types
                      );
  IF retval <= 0 THEN
#ifdef DEBUG
    IF (retval <> TCP_NOT_READY) | (timeout_ms > 0) THEN
      DEBUGLOG1("%010d-*** RecvSessionInfo: ReadCmdMsg(CMD_SESSINFO) failed, retval=%d", TO_UDINT(retval));
    END_IF;
#endif
    RETURN;
  END_IF;

  IF retval < (SIZEOF(msgSessInfo.cHdr.cmd) + SIZEOF(msgSessInfo.version) + SIZEOF(msgSessInfo.instId)) THEN
    // not enough data received !
    DEBUGLOG0("%010d-*** RecvSessionInfo: not enough data received");
    retval := ERR_INVALID_CMSGDATA;
    RETURN;
  END_IF;
  DEBUGLOG2("%010d-RecvSessionInfo: SESSINFO response received: version of peer=0x%08X, instId=0x%08X", cmsg$msgSessInfo.version, cmsg$msgSessInfo.instId);

  IF versionOfPeer <> NIL THEN
    versionOfPeer^ := cmsg$msgSessInfo.version;
    instIdOfPeer^  := cmsg$msgSessInfo.instId;

    IF retval >= (msgSessInfo.sizeofStatList + sizeof(msgSessInfo.sizeofStatList) - msgSessInfo.version) THEN
      sizeofRemoteDynList^  := cmsg$msgSessInfo.sizeofDynList;
      sizeofRemoteStatList^ := cmsg$msgSessInfo.sizeofStatList;
    END_IF;
  END_IF;

END_FUNCTION
#endif

//------------------------------------------------------------------------------
// ExchgSessionInfo
//
//  Exchange session info with the server
//------------------------------------------------------------------------------
#ifdef COMLINK_TCP_CLIENT
FUNCTION ExchgSessionInfo
VAR_INPUT
    bsock         : ^bufferedSocket;
    mySessId      : UDINT;
    timeout_ms    : UDINT;      // timeout, in milliseconds
    versionOfPeer : ^UDINT;
    instIdOfPeer  : ^UDINT;
    sizeofRemoteDynList  : ^UINT;
    sizeofRemoteStatList : ^UINT;
END_VAR
VAR_OUTPUT
    retval        : DINT;
END_VAR

  // Send the request
  retval := SendSessionInfo(bsock, mySessId, timeout_ms);
  IF retval <= 0 THEN
    RETURN;
  END_IF;

  // Read the response
  retval := RecvSessionInfo(bsock,
                            timeout_ms,
                            versionOfPeer,
                            instIdOfPeer,
                            sizeofRemoteDynList,
                            sizeofRemoteStatList
                            );
  IF retval <= 0 THEN
    RETURN;
  END_IF;

END_FUNCTION
#endif

#ifdef COMLINK_TCP_CLIENT
FUNCTION SetSocketOptions
VAR_INPUT
  sock : DINT;
END_VAR
VAR
  onOff : DINT;
END_VAR

  IF OS_TCP_USER_VERSION >= 5 THEN
   onOff := 0; // 0 means disable, 1 means enable
   OS_TCP_USER_SETSOCKOPT(sock, SOL_SOCKET, SO_DELAYED_ACK, #onOff$CHAR, sizeof(onOff));
   OS_TCP_USER_SETSOCKOPT(sock, SOL_SOCKET, SO_NAGLE,       #onOff$CHAR, sizeof(onOff));
  END_IF;

END_FUNCTION

FUNCTION CreateSocket
VAR_OUTPUT
  sock : DINT;
END_VAR

  sock := OS_TCP_USER_SOCKET();
  IF sock >= 0 THEN
    IF sock < arraysize(usedsocks) THEN
      usedsocks[sock] := 'L';
    END_IF;
    SetSocketOptions(sock);
  END_IF;

END_FUNCTION
#endif

//------------------------------------------------------------------------------
// CheckClientConnection
//
//  Check the connection from the client to the server and try to re-connect
//  when the connection does not exist.
//------------------------------------------------------------------------------
#ifdef COMLINK_TCP_CLIENT
FUNCTION CheckClientConnection
VAR_INPUT
    pLogin        : ^loginContext;  // connection context
    bsock         : ^bufferedSocket;
    timeout_ms    : UDINT;          // timeout, in milliseconds
END_VAR
VAR_OUTPUT
    retval        : comlinkReason;
END_VAR
VAR
    versionOfPeer : UDINT;
    instIdOfPeer  : UDINT;
    rc            : DINT;
    sizeofRemoteDynList  : UINT;
    sizeofRemoteStatList : UINT;
END_VAR

  IF bsock^.isInstIdVerified = INSTID_MISMATCH THEN
    // the server has been restarted, no retry possible
    retval := COMLINK_ERR_LOGIN_REQUIRED;
    RETURN;
  END_IF;

  IF (bsock^.sock >= 0) & (bsock^.isInstIdVerified = INSTID_MATCH) THEN
    // everything o.k., the connection is up and the server has not been restarted
    retval := COMLINK_OK;
    RETURN;
  END_IF;

  IF bsock^.sock < 0 THEN
    // the connection is down, start a reconnect process
    retval := COMLINK_ERR_NOCONNECTION;

    bsock^.isInstIdVerified := INSTID_NOT_VERIFIED;
    IF bsock^.pndSock >= 0 THEN
      // the socket is already in a 'connect pending' state
      RETURN;
    END_IF;

    bsock^.pndSock := CreateSocket();
    IF bsock^.pndSock < 0 THEN
      DEBUGLOG1("%010d-*** CheckClientConnection: CreateSocket failed, rc=%d", bsock^.pndSock$UDINT);
      RETURN;
    END_IF;

    // The connection is now in a 'connect pending' state. The CyWork task does the rest
    DEBUGLOG2("%010d-*** CheckClientConnection: connection is now in pending state (sock %d, pndSock %d)", bsock^.sock$UDINT, bsock^.pndSock$UDINT);
    RETURN;
  END_IF;

  // the connection is up, but the instance id of the server is not verified

  IF bsock^.isInstIdVerified = INSTID_NOT_VERIFIED THEN
    // send session information
    rc := SendSessionInfo(bsock, pLogin^.pComdefT$UDINT, timeout_ms);
    IF rc <= 0 THEN
      DEBUGLOG1("%010d-*** CheckClientConnection: SendSessionInfo failed, retval=%d", TO_UDINT(retval));
      CloseBufferedSock(bsock);
      RETURN;
    END_IF;
    bsock^.isInstIdVerified := INSTID_CMD_PENDING;
  END_IF;

  IF bsock^.isInstIdVerified = INSTID_CMD_PENDING THEN
    // receive session information
    sizeofRemoteDynList  := pLogin^.sizeofRemoteDynList;
    sizeofRemoteStatList := pLogin^.sizeofRemoteStatList;
    rc := RecvSessionInfo(bsock, timeout_ms, #versionOfPeer, #instIdOfPeer, #sizeofRemoteDynList, #sizeofRemoteStatList);
    IF rc <= 0 THEN
      IF (rc <> TCP_NOT_READY) | (timeout_ms > 0) THEN
        DEBUGLOG1("%010d-*** CheckClientConnection: RecvSessionInfo failed, retval=%d", TO_UDINT(retval));
        CloseBufferedSock(bsock);
      END_IF;
      RETURN;
    END_IF;
    IF pLogin^.instIdOfPeer = instIdOfPeer THEN
      DEBUGLOG0("%010d-CheckClientConnection: instance ID matches");
      pLogin^.sizeofRemoteDynList  := sizeofRemoteDynList;
      pLogin^.sizeofRemoteStatList := sizeofRemoteStatList;
      bsock^.isInstIdVerified := INSTID_MATCH;
    ELSE
      DEBUGLOG0("%010d-*** CheckClientConnection: instance ID does not match, closeing connection");
      bsock^.isInstIdVerified := INSTID_MISMATCH;
      CloseBufferedSock(bsock);
    END_IF;
  END_IF;

  IF bsock^.isInstIdVerified = INSTID_MATCH THEN
    retval := COMLINK_OK;
  ELSE
    retval := COMLINK_ERR_LOGIN_REQUIRED;
  END_IF;

END_FUNCTION
#endif

//------------------------------------------------------------------------------
// TraceMsg4Client
//------------------------------------------------------------------------------
FUNCTION TraceMsg4Client

  IF ComlinkT_wasTraceMsgDisplayed = 0 THEN

    IF isClientReady < 0 THEN
      CASE isClientReady OF
        COMLINKT_ERR_NOTCP:
          TRACE_ERR("Comlink/TCP client error: TCP_USER interface not available");
          LSLCLI_LoaderTracePrint("Comlink/TCP client error: TCP_USER interface not available", 12);
        COMLINKT_ERR_NOMTAPI:
          TRACE_ERR("Comlink/TCP client error: MT interface not available");
          LSLCLI_LoaderTracePrint("Comlink/TCP client error: MT interface not available", 12);
        COMLINKT_ERR_WRONG_OSVER:
          TRACE_ERR("Comlink/TCP client error: wrong OS-version (must be > 5.42)");
          LSLCLI_LoaderTracePrint("Comlink/TCP client error: wrong OS-version (must be > 5.42)", 12);
      ELSE
          TRACE_ERR("Comlink/TCP client error: unknown error code");
          LSLCLI_LoaderTracePrint("Comlink/TCP client error: unknown error code", 12);
      END_CASE;
      ComlinkT_wasTraceMsgDisplayed := 1;
      RETURN;
    END_IF;

  END_IF;

END_FUNCTION

FUNCTION TCPIP_Task
VAR_INPUT
  pvoid : ^void;
END_VAR;
//------------------------------------------------------------------------------
// ComlinkT_Init
//
//  Creates sockets for the command- and refresh- server and places them
//  into the listening state. The server queries its command port number from
//  the operating system. Usually it is port 1955, but when multiple servers
//  run on the same machine (e.g.LARS) then it can be a different number.
//  The refresh port number is the command port number plus 1.
//------------------------------------------------------------------------------
FUNCTION ComlinkT_Init
VAR
#ifdef COMLINK_TCP_SERVER
    cmdPortSrvr  : UDINT;
    refrPortSrvr : UDINT;
#endif
#ifdef COMLINK_TCP_CLIENT
    i            : UDINT;
#endif
END_VAR
  ComlinkT_wasTraceMsgDisplayed :=0;
#ifdef COMLINK_TCP_SERVER
  isServerReady     := COMLINKT_ERR_NOTCP;
  pCmdConnRoot      := NIL;
  pRefrConnRoot     := NIL;
  nbrCmdConn        := 0;
  nbrRefrConn       := 0;
  nbrRecycled       := 0;
  pRefrConnDataRoot := NIL;
  tcpServerState    := 0;
  tcpAcceptState    := 0;
  s_pCmdConn        := NIL;
  s_pRefrConn       := NIL;

#endif
#ifdef COMLINK_TCP_CLIENT
  isClientReady     := COMLINKT_ERR_NOTCP;
  FOR i := 0 TO (g_max_logins - 1) DO
    loginArray[i] := NIL;
  END_FOR;
  loginAnz          := 0;
  g_pCallback       := NIL;
#ifdef LOADER_TCP_MODERATE
  //SCHMAT_001
  TCPCltCntr        := 0;
#endif
#endif
  myInstanceId      := GetMyInstanceId();
  myApplId          := GetMyApplId();

  IF OS_CILGET("TCP_USER", #lsl_tcp_user) THEN
    // the OS does not support TCP/IP
    DEBUGLOG0("%010d-TCP_USER interface not supported");
    lsl_tcp_user  := NIL;
    #ifdef COMLINK_TCP_SERVER
    cmdSockSrvr   := INVALID_SOCKET_NUM;
    refrSockSrvr  := INVALID_SOCKET_NUM;
    #endif
    RETURN;
  END_IF;

#ifdef COMLINK_TCP_CLIENT
  isClientReady := 0;
  IF mt_api = NIL THEN
    DEBUGLOG0("%010d-LSL_MULTITASK interface not supported");
    isClientReady := COMLINKT_ERR_NOMTAPI;
  END_IF;

  IF _RtOSversion < 16#052B THEN
      // there was a bug with LSL_MULTITASK in OS <= 5.42
    isClientReady     := COMLINKT_ERR_WRONG_OSVER;
  END_IF;

  loginArrayMutex := OS_MT_CreateSemaphore(MTSEMATYPE_MUTEX,
                                           1,    // initvalue
                                           0,    // flags: 0 means create unconitionally
                                           "COMLINKT0"
                                           );
  IF loginArrayMutex = NIL THEN
    isClientReady := COMLINKT_ERR_API_FAILED;
  END_IF;

#endif

#ifdef COMLINK_TCP_SERVER
  isServerReady := 0;
  cmdPortSrvr := 0;
  IF lsl_tcp_user^.udVersion >= 3 THEN
    cmdPortSrvr := OS_TCP_USER_GETSERVBYNAME("comlink", "tcp");
  END_IF;
  IF cmdPortSrvr = 0 THEN
    cmdPortSrvr  := 1955;               // default cmd port is hardcoded to 1955
  END_IF;
  refrPortSrvr := cmdPortSrvr + 1;

  cmdSockSrvr  := CreateSocket(); // create a new command socket
  refrSockSrvr := CreateSocket(); // create a new refresh socket

  IF (cmdSockSrvr >= 0) & (refrSockSrvr >= 0) THEN
    // place the sockets into the listening state
    IF OS_TCP_USER_LISTEN(cmdSockSrvr, cmdPortSrvr, 0) <> TCP_NO_ERROR THEN
      DEBUGLOG0("%010d-TCP Server for command data not started");
      TRACE_ERR("TCP Server for command data not started");
      LSLCLI_LoaderTracePrint("TCP Server for command data not started", 12);
      isServerReady := COMLINKT_ERR_API_FAILED;
    ELSE
      IF OS_TCP_USER_LISTEN(refrSockSrvr, refrPortSrvr, 0) <> TCP_NO_ERROR THEN
        DEBUGLOG0("%010d-TCP Server for refresh data not started");
        TRACE_ERR("TCP Server for refresh data not started");
        LSLCLI_LoaderTracePrint("TCP Server for refresh data not started", 12);
        isServerReady := COMLINKT_ERR_API_FAILED;
      ELSE
        // everything o.k.
        DEBUGLOG2("%010d-ComlinkT_Init:server started, cmdPort=%d, refrPort=%d", cmdPortSrvr$UDINT, refrPortSrvr$UDINT);
      END_IF;
    END_IF;
  ELSE
    isServerReady := COMLINKT_ERR_API_FAILED;
  END_IF;

  IF isServerReady < 0 THEN
    // something was wrong, cleanup now
    DEBUGLOG0("%010d-*** ComlinkT_Init:server did not start");
    IF cmdSockSrvr >= 0 THEN
      CloseSock(#cmdSockSrvr);
    END_IF;
    IF refrSockSrvr >= 0 THEN
      CloseSock(#refrSockSrvr);
    END_IF;
  END_IF;
#endif

#ifdef LOADER_TCP_MODERATE
  taskhandle := OS_MT_CREATETHREAD(#TCPIP_Task(),
                                   14,
                                   16#4000,
                                   MT_Task_SAVETHIS,
                                   NIL,
                                   "LDR_TCPIP_Task");

  //udTimeTCP := 0;
#endif
END_FUNCTION
//------------------------------------------------------------------------------
// ComlinkT_Login
//
//  Establish a connection to a comlink server.
//------------------------------------------------------------------------------
#ifdef COMLINK_TCP_CLIENT
FUNCTION ComlinkT_Login
VAR_INPUT
    pComdef       : ^comdef;
END_VAR
VAR_OUTPUT
    retval        : UINT;
END_VAR
VAR
    pComdefT      : ^comdefT;
    pLogin        : ^loginContext; // connection context
    cmdPortSrvr   : UDINT;        // port number of the servers command port
    refrPortSrvr  : UDINT;        // port number of the servers refresh port
    versionOfPeer : UDINT;
    instIdOfPeer  : UDINT;
    rc            : DINT;
    i             : UDINT;
    sizeofRemoteDynList  : UINT;
    sizeofRemoteStatList : UINT;
END_VAR

  pComdefT := pComdef$^comdefT;
  retval   := COMLINK_ERR_GENERAL;

  DEBUGLOG1("%010d-ComlinkT_Login: ip-address=0x%08X", pComdefT^.ipAddress$UDINT);

  IF isClientReady < 0 THEN
    DEBUGLOG0("%010d-*** ComlinkT_Login: client is not ready");
    TraceMsg4Client();
    retval := COMLINK_ERR_CLIENT_NOTREADY;
    RETURN;
  END_IF;

  IF (pComdefT^.interface <> IF_TYPE_TCPIP1) &
     (pComdefT^.interface <> IF_TYPE_TCPIP1_NEW) THEN
    // no other interface type than TCPIP1 is supported in the moment.
    DEBUGLOG0("%010d-*** ComlinkT_Login: invalid interface type");
    retval := COMLINK_ERR_UNSUPPORTED_INTERFACE;
    RETURN;
  END_IF;

  IF (pComdefT^.interface = IF_TYPE_TCPIP1_NEW) & (pComdefT^.port <> 0) THEN
    cmdPortSrvr  := pComdefT^.port;
  ELSE
    cmdPortSrvr  := 1955;
  END_IF;
  refrPortSrvr := cmdPortSrvr + 1;

  // try to get a connection context
  pLogin := AllocateLoginContext(pComdefT^.ipAddress, cmdPortSrvr);
  IF pLogin = NIL THEN
    DEBUGLOG0("%010d-*** ComlinkT_Login: AllocateLoginContext failed");
    RETURN;
  END_IF;

  // establish a connection to the command server
  pLogin^.cmdSockClnt.sock := CreateSocket();
  IF pLogin^.cmdSockClnt.sock < 0 THEN
    DEBUGLOG1("%010d-*** ComlinkT_Login: CreateSocket failed, rc=%d", pLogin^.cmdSockClnt.sock$UDINT);
    GOTO EndLabel;
  END_IF;
  rc := Connect(pLogin^.cmdSockClnt.sock,
                pLogin^.ipAddrSrvr,
                cmdPortSrvr,
                CLIENT_TIMEOUT_CONNECT
                );
  IF rc < 0 THEN
    DEBUGLOG1("%010d-*** ComlinkT_Login: Connect to command server failed, rc=%d", TO_UDINT(rc));
    retval := COMLINK_ERR_NOCONNECTION;
    GOTO EndLabel;
  END_IF;
  DEBUGLOG2("%010d-ComlinkT_Login: connected to command server (port:%d, sock%d)", cmdPortSrvr$UDINT, pLogin^.cmdSockClnt.sock$UDINT);

  // establish a connection to the refresh server
  pLogin^.refrSockClnt.sock := CreateSocket();
  IF pLogin^.refrSockClnt.sock < 0 THEN
    DEBUGLOG1("%010d-*** ComlinkT_Login: CreateSocket failed, rc=%d", pLogin^.refrSockClnt.sock$UDINT);
    GOTO EndLabel;
  END_IF;
  rc := Connect(pLogin^.refrSockClnt.sock,
                pLogin^.ipAddrSrvr,
                refrPortSrvr,
                CLIENT_TIMEOUT_CONNECT
                );
  IF rc < 0 THEN
    DEBUGLOG1("%010d-*** ComlinkT_Login: Connect to refresh server failed, rc=%d", TO_UDINT(rc));
    retval := COMLINK_ERR_NOCONNECTION;
    GOTO EndLabel;
  END_IF;
  DEBUGLOG2("%010d-ComlinkT_Login: connected to refresh server (port:%d, sock%d)", refrPortSrvr$UDINT, pLogin^.refrSockClnt.sock$UDINT);

  // exchange session info with the server
  sizeofRemoteDynList  := pLogin^.sizeofRemoteDynList;
  sizeofRemoteStatList := pLogin^.sizeofRemoteStatList;
  rc := ExchgSessionInfo(#pLogin^.refrSockClnt,
                         pComdef$UDINT,
                         CLIENT_TIMEOUT_REQ,
                         #versionOfPeer,
                         #instIdOfPeer,
                         #sizeofRemoteDynList,
                         #sizeofRemoteStatList);
  IF rc <= 0 THEN
    DEBUGLOG2("%010d-*** ComlinkT_Login(sock %d): ExchgSessionInfo failed, rc=%d", pLogin^.refrSockClnt$UDINT, TO_UDINT(rc));
    retval := COMLINK_ERR_NOCONNECTION;
    GOTO EndLabel;
  END_IF;

  retval := 0;
  pLogin^.versionOfPeer := versionOfPeer;
  pLogin^.instIdOfPeer  := instIdOfPeer;
  pLogin^.sizeofRemoteDynList  := sizeofRemoteDynList;
  pLogin^.sizeofRemoteStatList := sizeofRemoteStatList;
  pLogin^.pComdefT      := pComdefT; // this pointer is needed when the callback function is called
  pLogin^.cmdSockClnt.isInstIdVerified  := INSTID_MATCH;
  pLogin^.refrSockClnt.isInstIdVerified := INSTID_MATCH;

  // Die SessionInfo wird jetzt auch über die CmdConn geschickt, damit der Server die Chance
  // hat inaktive CmdConns zu erkennen und freizugeben. Der Returncode wird nicht ausgewertet,
  // das es alte Loaderversionen geben kann, die auf der CmdConn den SessionInfo Befehl nicht
  // verstehen.
  ExchgSessionInfo(#pLogin^.cmdSockClnt, pComdef$UDINT, CLIENT_TIMEOUT_REQ, NIL, NIL, NIL, NIL);

EndLabel:
  IF retval <> 0 THEN
    // something was wrong, cleanup now
    ReleaseLoginContext(pLogin);
  ELSE
    // success: try to put pLogin into loginArray
    OS_MT_Wait(loginArrayMutex);

    // search for a connection context already in use
    FOR i := 0 TO (g_max_logins - 1) DO
      IF loginArray[i] <> NIL THEN
        IF (loginArray[i]^.ipAddrSrvr = pLogin^.ipAddrSrvr) &
           (loginArray[i]^.cmdPortSrvr = pLogin^.cmdPortSrvr) THEN
          // address is already in use
          IF loginArray[i]^.pComdefT = pComdefT THEN
            // gleiches pcomdef bedeutet reconnect -> das bisgherige pcomdef wird daher freigegeben
            (*
               In ReleaseLoginContext (aus UnlockLoginContext aufgerufen, falls refCnt 0 ist),
               wird pLogin^.pComdefT^.pLogin auf NIL gesetzt wird, falls pLogin^.pComdefT <> NIL ist.
               Es soll damit verhindert werden, dass in der pComdefT Struktur, die ja vom
               Aufrufer bereitgestellt wird, ein Verweis auf die freigegebene Login-Struktur
               existiert. Weiter unten wird dann pComdefT^.pLogin auf die neue Login-Struktur gesetzt.

               Hier könnte es zu einem Fehler kommen, wenn ReleaseLoginContext in diesem
               UnlockLoginContext noch nicht aufgerufen wird, weil der RefCnt > 0 ist.
               Das kann passieren, wenn der ComlinkT_Login Aufruf aus dem Background erfolgt,
               während im Cyclic gerade der Login-Context gelockt ist (ComlinkT_CyWork_Client).
               Wenn dann ReleaseLoginContext aufgerufen wird, nachdem weiter unten pComdefT^.pLogin
               auf den neuen Wert gesetzt wurde, dann wird pComdefT^.pLogin in ReleaseLoginContext
               wieder auf 0 gesetzt.

               Um das zu verhindern, wird hier die Referenz auf die Comdef Struktur des Aufrufers
               auf NIL gesetzt.
            *)
            loginArray[i]^.pComdefT := NIL;
            UnlockLoginContext(loginArray[i]);
            EXIT;
          END_IF;
          // bei ungleichem pcomdef wird ein neuer channel aufgemacht (vor 2.6 wurde ADDR_IN_USE zurückgegeben)
        END_IF;
      END_IF;
    END_FOR;

    // search a free entry in loginArray
    FOR i := 0 TO (g_max_logins - 1) DO
      IF loginArray[i] = NIL THEN
        EXIT;
      END_IF;
    END_FOR;
    IF i = g_max_logins THEN
      retval := COMLINK_ERR_MAXCONN;
      OS_MT_Signal(loginArrayMutex);
      ReleaseLoginContext(pLogin);
      RETURN;
    END_IF;

    pComdefT^.pLogin := pLogin;
    // make an entry in the loginArray
    loginArray[i] := pLogin;
    loginAnz += 1;

    OS_MT_Signal(loginArrayMutex);
  END_IF ;

END_FUNCTION
#endif

//------------------------------------------------------------------------------
// ComlinkT_Logout
//
//  Close a connection to a comlink server.
//------------------------------------------------------------------------------
#ifdef COMLINK_TCP_CLIENT
FUNCTION ComlinkT_Logout
VAR_INPUT
    pComdef       : ^comdef;
END_VAR
VAR
    pComdefT      : ^comdefT;
    pLogin        : ^loginContext; // connection context
    startTime     : udint;
END_VAR

  pComdefT := pComdef$^comdefT;

  IF isClientReady < 0 THEN
    DEBUGLOG0("%010d-*** ComlinkT_Logout: client is not ready");
    TraceMsg4Client();
    RETURN;
  END_IF;

  pLogin := pComdefT^.pLogin;
  IF pLogin = NIL THEN
    RETURN;
  END_IF;
  IF pLogin^.instIdOfPeer = 0x1AFEE THEN
    // es hat bereits ein Logout stattgefunden
    RETURN;
  END_IF;
  // Da instIdOfPeer ab jetzt nicht mehr benötigt wird, wird der Magic Value 0x1AFEE
  // in instIdOfPeer dafür verwendet, einen doppelten Logout Aufruf zu erkennen.
  pLogin^.instIdOfPeer := 0x1AFEE;

  LockLoginContext2(pLogin);

  SendLogout( pComdefT );

  // 20ms nach dem Senden des Logout warten
  startTime := ops.tAbsolute;
  WHILE (ops.tAbsolute - startTime) < 20 DO
    OS_MT_Delay(1);
  END_WHILE;

  UnlockLoginContext(pLogin); // wg. dem LockLoginContext2 Aufruf in dieser Funktion
  UnlockLoginContext(pLogin); // wg. dem LockLoginContext im ComlinkT_Login

END_FUNCTION
#endif

//------------------------------------------------------------------------------
// ComlinkT_TxCommandEx
//
//  This function send interpreter code to the comlink server. The server
//  executes the code and responds with the the result and the workstate.
//------------------------------------------------------------------------------
#ifdef COMLINK_TCP_CLIENT
FUNCTION ComlinkT_TxCommandEx
VAR_INPUT
    opCode    : UDINT;
    length    : UDINT;
    aPara     : ^USINT;
    pComdef   : ^comdef;
    pResu     : ^UDINT;
    pStatus   : ^IPRSTATES;
    res       : UDINT;
END_VAR
VAR_OUTPUT
    retval    : comlinkReason;
END_VAR
VAR
    pComdefT  : ^comdefT;
    pLogin    : ^loginContext; // connection context
    reqMsg    : msgBefiprReq; // request structure for command CMD_BEFIPR
    reqMsgLen : UDINT;
    fOk       : UDINT;
    ack       : UDINT;
    rc        : DINT;
    rc2       : comlinkReason;
END_VAR

  pComdefT := pComdef$^comdefT;
  pStatus^ := ERROR;
  retval   := COMLINK_ERR_GENERAL;
  fOk   := 0;

  IF isClientReady < 0 THEN
    DEBUGLOG0("%010d-*** ComlinkT_TxCommandEx: client is not ready");
    TraceMsg4Client();
    retval := COMLINK_ERR_CLIENT_NOTREADY;
    RETURN;
  END_IF;

  pLogin := pComdefT^.pLogin;
  IF pLogin = NIL THEN
    retval := COMLINK_ERR_LOGIN_REQUIRED;
    RETURN;
  END_IF;
  LockLoginContext2(pLogin);

  rc2 := CheckClientConnection(pLogin, #pLogin^.cmdSockClnt, CLIENT_TIMEOUT_REQ);
  IF rc2 <> COMLINK_OK THEN
    retval := rc2;
    UnlockLoginContext(pLogin); // wg. dem LockLoginContext2 Aufruf in dieser Funktion
    RETURN;
  END_IF;

  pResu^ := (#pLogin^.befiprResp.resu)$UDINT;

  IF pLogin^.cmdSockClnt.sock < 0 THEN
    // no connection exists
    DEBUGLOG0("%010d-*** ComlinkT_TxCommandEx: no connection exists");
    retval := COMLINK_ERR_NOCONNECTION;
    UnlockLoginContext(pLogin); // wg. dem LockLoginContext2 Aufruf in dieser Funktion
    RETURN;
  END_IF;

  IF length > SIZEOF(reqMsg.instr.aPara) THEN
    // parameter length is too big
    DEBUGLOG0("%010d-*** ComlinkT_TxCommandEx: parameter length is too big");
    retval := COMLINK_ERR_INVALID_PARAM;
    UnlockLoginContext(pLogin); // wg. dem LockLoginContext2 Aufruf in dieser Funktion
    RETURN;
  END_IF;

  // prepare the request message structure
  reqMsg.workState    := BUSY;
  reqMsg.instr.opCode := opCode$INSTRSET;
  reqMsg.instr.uiLng  := (length + SIZEOF(instruct.uiLng))$UINT;
  _memcpy(#reqMsg.instr.aPara, aPara, length);

  reqMsgLen := SIZEOF(cmdMsgHdr)           +
               SIZEOF(reqMsg.workState)    +
               SIZEOF(reqMsg.instr.opCode) +
               SIZEOF(reqMsg.instr.uiLng)  +
               length;

  // Send the request
  rc := SendCmdMsg(#pLogin^.cmdSockClnt,
                   CMD_BEFIPR,
                   MASK_CMD_ACK,      // Type and Ack field of command (type: request, ack: a response is required)
                   #reqMsg$cMessage,
                   reqMsgLen,
                   CLIENT_TIMEOUT_REQ,
                   0,                 // do not use buffered sends
                   0                  // fFlush
                  );
  IF rc <= 0 THEN
    DEBUGLOG1("%010d-*** ComlinkT_TxCommandEx: SendCmdMsg failed, rc=%d", TO_UDINT(rc));
    retval := COMLINK_ERR_NOCONNECTION;
    GOTO EndLabel;
  END_IF;
  DEBUG_VERBOSE2("%010d-ComlinkT_TxCommandEx: BEFIPR request sent, opCode=%d, msgLen=%d", opCode, TO_UDINT(rc));

  // Read the response
  rc := ReadCmdMsg(#pLogin^.cmdSockClnt,
                   #pLogin^.befiprResp$cMessage,
                   SIZEOF(pLogin^.befiprResp),
                   CLIENT_TIMEOUT_REQ,
                   #ack,                // received ack field
                   CMD_BEFIPR,
                   CMD_TYPE_RESP        // accept only response types
                  );
  IF rc <= 0 THEN
    DEBUGLOG1("%010d-*** ComlinkT_TxCommandEx: ReadCmdMsg failed, rc=%d", TO_UDINT(rc));
    retval := COMLINK_ERR_NOCONNECTION;
    GOTO EndLabel;
  END_IF;
  AliveCheckMsgRcvd(pLogin);

  IF rc < (SIZEOF(pLogin^.befiprResp.cHdr.cmd) + SIZEOF(pLogin^.befiprResp.workstate)) THEN
    // not enough data received !
    DEBUGLOG0("%010d-*** ComlinkT_TxCommandEx: not enough data received");
    retval := COMLINK_ERR_INVALID_RESPONSE;
    GOTO EndLabel;
  END_IF;

  fOk := 1;

EndLabel:
  IF fOk = 0 THEN
    // The connection has to be closed because it's possible that partial data
    // is transferred.
    DEBUGLOG0("%010d-ComlinkT_TxCommandEx: closing socket");
    CloseBufferedSock(#pLogin^.cmdSockClnt);
    pStatus^ := ERROR;
  ELSE
    IF ack THEN
      pStatus^ := pLogin^.befiprResp.workstate;
      DEBUG_VERBOSE2("%010d-ComlinkT_TxCommandEx: BEFIPR response received, dataLen=%d, Status=%d", TO_UDINT(rc-4), pStatus^$UDINT);
      //DEBUG_VERBOSE3("%010d-                    uiLng=%d, aData[0]=0x%08X, aData[4]=0x%08X", TO_UDINT(pLogin^.befiprResp.resu.uiLng), pLogin^.befiprResp.resu.aData[0]$UDINT, pLogin^.befiprResp.resu.aData[4]$UDINT);
      retval := COMLINK_IPR;
    ELSE
      pStatus^ := ERROR;
      DEBUGLOG0("%010d-ComlinkT_TxCommandEx: NACK received");
      retval := COMLINK_ERR_INVALID_RESPONSE;
    END_IF;
  END_IF;
  UnlockLoginContext(pLogin); // wg. dem LockLoginContext2 Aufruf in dieser Funktion

END_FUNCTION
#endif

//------------------------------------------------------------------------------
// ComlinkT_TxUpd_nocs
//------------------------------------------------------------------------------
#ifdef COMLINK_TCP_CLIENT
FUNCTION ComlinkT_TxUpd_nocs
VAR_INPUT
    pLslcommregdata : ^lslCommregData;
    pLogin          : ^loginContext; // connection context
    uiflags         : UINT;
END_VAR
VAR_OUTPUT
    retval          : comlinkReason;
END_VAR
VAR
    reqMsg        : msgTxUpdReq;   // request structure for command CMD_TXUPD
    pt_comStCell  : ^comStCell;
    timeout_ms    : UDINT;         // timeout value for send request
    fFlush        : UDINT;
    updList       : ^updateList;
    listIndex     : UDINT;
    listType      : UDINT;
    rc            : DINT;
    rc2           : comlinkReason;
    timx          : udint;
END_VAR

  retval := COMLINK_ERR_GENERAL;

  rc2 := CheckClientConnection(pLogin, #pLogin^.refrSockClnt, 0);
  IF rc2 <> COMLINK_OK THEN
    retval := rc2;
    RETURN;
  END_IF;

  IF pLslcommregdata^.varpos$INT < 1000 THEN
    updList   := #pLogin^.statList;
    listIndex := pLslcommregdata^.varpos;
    listType  := 0;
  ELSE
    updList   := #pLogin^.dynList;
    listIndex := pLslcommregdata^.varpos - 1000;
    listType  := 1;
  END_IF;

  IF listIndex >= updList^.nbrCells THEN
    IF IncreaseUpdateList(updList, listIndex + 1, listType) = NIL THEN
      DEBUGLOG0("%010d-*** ComlinkT_TxUpd: MemoryUpdateList failed");
      CloseBufferedSock(#pLogin^.refrSockClnt);
      RETURN;
    END_IF;
    DEBUGLOG2("%010d-*** ComlinkT_TxUpd: list %d increased to %d entries", listType, updList^.nbrCells);
  END_IF;

  pt_comStCell := updList^.pFirstCell + (listIndex * SIZEOF (comStCell));

  timx                       := pLslcommregdata^.uiTime; // u32 := u16
  pt_comStCell^.dData        := 16#80000001$DINT;     // INVALID
  pt_comStCell^.pCh          := pLslcommregdata^.LASALID$^SVRCH;
  pt_comStCell^.udUpdateRate := (timx and 16#3FFF) or ((timx and 16#C000) shl 16) or (uiflags shl 14);
  pt_comStCell^.udUpdateRate := pt_comStCell^.udUpdateRate or UPDRATE_FLAG_FORCE_CHANGE;
  pt_comStCell^.VarlistID    := pLslcommregdata^.VarlistID;
  pt_comStCell^.udLastUpdate := 0;

  // prepare the request message structure
  reqMsg.iOff    := pLslcommregdata^.varpos$UINT;
  reqMsg.comcell := pt_comStCell^;  // copy struct on struct;

  IF QUERY_FREE_TXBUF(pLogin^.refrSockClnt) < (2 * SIZEOF(reqMsg)) THEN
    DEBUGLOG0("%010d-*** ComlinkT_TxUpd: send buffer shortage, next send will block");
    timeout_ms := CLIENT_TIMEOUT_REQ;
    fFlush := 1;
  ELSE
    timeout_ms := 0;    // timeout: non-blocking
    fFlush := 0;
  END_IF;

  // Send the request
  rc := SendCmdMsg(#pLogin^.refrSockClnt,
                   CMD_TXUPD,
                   0,                // Type and Ack field of command (type: request, ack: no response required)
                   #reqMsg$cMessage,
                   SIZEOF(reqMsg),
                   timeout_ms,
                   1,                // use bufferd send
                   fFlush            // fFlush
                  );
  IF rc <= 0 THEN
    DEBUGLOG2("%010d-*** ComlinkT_TxUpd(VarPos %d): SendCmdMsg failed, rc=%d", pLslcommregdata^.varpos, TO_UDINT(rc));
    CloseBufferedSock(#pLogin^.refrSockClnt);
    retval := COMLINK_ERR_NOCONNECTION;
  ELSE
    DEBUG_VERBOSE3("%010d-ComlinkT_TxUpd: TXUPD request sent, msgLen=%d, VarPos=%d, time=0x%08X", TO_UDINT(rc), TO_UDINT(pLslcommregdata^.varpos), TO_UDINT(pLslcommregdata^.uiTime));
    retval := COMLINK_OK;
  END_IF;

END_FUNCTION
#endif

//------------------------------------------------------------------------------
// ComlinkT_TxUpd
//
// Return value:
//  If the function succeeds, the return value is 0, othzerwise it is a
//  negative error code.
//------------------------------------------------------------------------------
#ifdef COMLINK_TCP_CLIENT
FUNCTION ComlinkT_TxUpd
VAR_INPUT
    pLslcommregdata : ^lslCommregData;
    pComdef         : ^comdef;
    res             : UDINT;
    uiflags         : UINT;
END_VAR
VAR_OUTPUT
    retval          : comlinkReason;
END_VAR
VAR
    pLogin          : ^loginContext; // connection context
END_VAR

  IF isClientReady < 0 THEN
    DEBUGLOG0("%010d-*** ComlinkT_TxUpd: client is not ready");
    TraceMsg4Client();
    retval := COMLINK_ERR_CLIENT_NOTREADY;
    RETURN;
  END_IF;

  pLogin := pComdef^$comdefT.pLogin;
  IF pLogin = NIL THEN
    retval := COMLINK_ERR_LOGIN_REQUIRED;
    RETURN;
  END_IF;

  OS_MT_Wait(pLogin^.hMutex);
  retval := ComlinkT_TxUpd_nocs(pLslcommregdata, pLogin, uiflags);
  OS_MT_Signal(pLogin^.hMutex);

END_FUNCTION
#endif

//------------------------------------------------------------------------------
// SendMaxIdleTime_TCP_nocs
//------------------------------------------------------------------------------
#ifdef COMLINK_TCP_CLIENT
FUNCTION SendMaxIdleTime_TCP_nocs
VAR_INPUT
  pComdefT : ^comdefT;
  remoteMaxIdleTime_ms : UDINT;
  pLogin          : ^loginContext; // connection context
END_VAR
VAR_OUTPUT
  retVal : DINT;
END_VAR
VAR
    reqMsg        : msgIdlTimReq;  // request structure for command CMD_MAXIDLETIME
    timeout_ms    : UDINT;         // timeout value for send request
    fFlush        : UDINT;
    rc            : DINT;
    rc2           : comlinkReason;
END_VAR

  retval := COMLINK_ERR_GENERAL;

  rc2 := CheckClientConnection(pLogin, #pLogin^.refrSockClnt, 0);
  IF rc2 <> COMLINK_OK THEN
    retval := rc2;
    RETURN;
  END_IF;

  // prepare the request message structure
  reqMsg.maxIdleTime_ms := remoteMaxIdleTime_ms;

  IF QUERY_FREE_TXBUF(pLogin^.refrSockClnt) < (2 * SIZEOF(reqMsg)) THEN
    DEBUGLOG0("%010d-*** SendMaxIdleTime_TCP_nots: send buffer shortage, next send will block");
    timeout_ms := CLIENT_TIMEOUT_REQ;
    fFlush := 1;
  ELSE
    timeout_ms := 0;    // timeout: non-blocking
    fFlush := 0;
  END_IF;

  // Send the request
  rc := SendCmdMsg(#pLogin^.refrSockClnt,
                   CMD_MAXIDLETIME,
                   0,                // Type and Ack field of command (type: request, ack: no response required)
                   #reqMsg$cMessage,
                   SIZEOF(reqMsg),
                   timeout_ms,
                   1,                // use bufferd send
                   fFlush            // fFlush
                  );
  IF rc <= 0 THEN
    DEBUGLOG1("%010d-*** SendMaxIdleTime_TCP_nots: SendCmdMsg failed, rc=%d", TO_UDINT(rc));
    CloseBufferedSock(#pLogin^.refrSockClnt);
    retval := COMLINK_ERR_NOCONNECTION;
  ELSE
    DEBUG_VERBOSE0("%010d-SendMaxIdleTime_TCP_nots: MAXIDLETIME request sent");
    retval := COMLINK_OK;
  END_IF;

END_FUNCTION

FUNCTION SendLOGOUT_TCP_nocs
VAR_INPUT
  pComdefT : ^comdefT;
  pLogin          : ^loginContext; // connection context
END_VAR
VAR_OUTPUT
  retVal : DINT;
END_VAR
VAR
    reqLOGOUT     : msgLOGOUTReq;
    rc            : DINT;
    rc2           : comlinkReason;
END_VAR

  retval := COMLINK_ERR_GENERAL;

  rc2 := CheckClientConnection(pLogin, #pLogin^.refrSockClnt, 0);
  IF rc2 <> COMLINK_OK THEN
    retval := rc2;
    RETURN;
  END_IF;

  rc := SendCmdMsg(#pLogin^.refrSockClnt,
                   CMD_LOGOUT,
                   0,      // Type and Ack field of command (type: request, ack: a response is required)
                   #reqLOGOUT$cMessage,
                   SIZEOF(reqLOGOUT),
                   10000,
                   1,                 // use buffered sends
                   1                  // fFlush
                  );

  IF rc <= 0 THEN
    DEBUGLOG1("%010d-*** SendLOGOUT_TCP_nots: SendCmdMsg failed, rc=%d", TO_UDINT(rc));
    CloseBufferedSock(#pLogin^.refrSockClnt);
    retval := COMLINK_ERR_NOCONNECTION;
  ELSE
    DEBUG_VERBOSE0("%010d-SendLOGOUT_TCP_nots: LOGOUT request sent");
    retval := COMLINK_OK;
    FLUSH_TXBUF( #pLogin^.refrSockClnt ); //safety
  END_IF;

  rc := SendCmdMsg(#pLogin^.cmdSockClnt,
                   CMD_LOGOUT,
                   0,      // Type and Ack field of command (type: request, ack: a response is required)
                   #reqLOGOUT$cMessage,
                   SIZEOF(reqLOGOUT),
                   10000,
                   1,                 // use buffered sends
                   1                  // fFlush
                  );

  IF rc <= 0 THEN
    DEBUGLOG1("%010d-*** SendLOGOUT_TCP_nots: SendCmdMsg failed, rc=%d", TO_UDINT(rc));
    CloseBufferedSock(#pLogin^.cmdSockClnt);
    retval := COMLINK_ERR_NOCONNECTION;
  ELSE
    DEBUG_VERBOSE0("%010d-SendLOGOUT_TCP_nots: LOGOUT request sent");
    retval := COMLINK_OK;
    FLUSH_TXBUF( #pLogin^.cmdSockClnt ); //safety
  END_IF;

END_FUNCTION

#endif

//------------------------------------------------------------------------------
// SendMaxIdleTime_TCP
//
// Return value:
//  If the function succeeds, the return value is 0, othzerwise it is a
//  negative error code.
//------------------------------------------------------------------------------
#ifdef COMLINK_TCP_CLIENT
FUNCTION SendMaxIdleTime_TCP
VAR_INPUT
  pComdefT : ^comdefT;
  remoteMaxIdleTime_ms : UDINT;
END_VAR
VAR_OUTPUT
  retVal : DINT;
END_VAR
VAR
    pLogin          : ^loginContext; // connection context
END_VAR

  IF isClientReady < 0 THEN
    DEBUGLOG0("%010d-*** ComlinkT_TxUpd: client is not ready");
    TraceMsg4Client();
    retval := COMLINK_ERR_CLIENT_NOTREADY;
    RETURN;
  END_IF;

  pLogin := pComdefT^.pLogin;
  IF pLogin = NIL THEN
    retval := COMLINK_ERR_LOGIN_REQUIRED;
    RETURN;
  END_IF;
  LockLoginContext2(pLogin);

  OS_MT_Wait(pLogin^.hMutex);
  retval := SendMaxIdleTime_TCP_nocs(pComdefT, remoteMaxIdleTime_ms, pLogin);
  OS_MT_Signal(pLogin^.hMutex);

  UnlockLoginContext(pLogin); // wg. dem LockLoginContext2 Aufruf in dieser Funktion

END_FUNCTION
#endif

#ifdef COMLINK_TCP_CLIENT
FUNCTION SendLogout_TCP
VAR_INPUT
  pComdefT : ^comdefT;
END_VAR
VAR_OUTPUT
  retVal : DINT;
END_VAR
VAR
    pLogin          : ^loginContext; // connection context
END_VAR

  IF isClientReady < 0 THEN
    DEBUGLOG0("%010d-*** ComlinkT_TxUpd: client is not ready");
    TraceMsg4Client();
    retval := COMLINK_ERR_CLIENT_NOTREADY;
    RETURN;
  END_IF;

  pLogin := pComdefT^.pLogin;
  IF pLogin = NIL THEN
    retval := COMLINK_ERR_LOGIN_REQUIRED;
    RETURN;
  END_IF;
  LockLoginContext2(pLogin);
